// TIA Portal V19 export
FUNCTION_BLOCK "ALL_AI"   // FB3, FBD
{ S7_Optimized_Access := 'TRUE' }
// stored: MemoryReserve 100, SetENOAutomatically false
   VAR
      AI_TT01 { S7_SetPoint := 'True'} : "AI";
      AI_TT02 { S7_SetPoint := 'True'} : "AI";
      AI_TT03 { S7_SetPoint := 'True'} : "AI";
      AI_CHS_TT01 { S7_SetPoint := 'True'} : "AI";
      AI_CHS_TT02 { S7_SetPoint := 'True'} : "AI";
      AI_CHS_TT03 { S7_SetPoint := 'True'} : "AI";
      AI_CHS_TT04 { S7_SetPoint := 'True'} : "AI";
      AI_CHS_MGLT { S7_SetPoint := 'True'} : "AI";
      AI_R2_TT01 { S7_SetPoint := 'True'} : "AI";
      AI_R2_TT02 { S7_SetPoint := 'True'} : "AI";
      AI_R2_TT03 { S7_SetPoint := 'True'} : "AI";
      AI_R3_TT01 { S7_SetPoint := 'True'} : "AI";
      AI_R3_TT02 { S7_SetPoint := 'True'} : "AI";
      AI_R3_TT03 { S7_SetPoint := 'True'} : "AI";
      AI_R4_TT03 { S7_SetPoint := 'True'} : "AI";
      AI_R4_TT02 { S7_SetPoint := 'True'} : "AI";
      AI_R4_TT01 { S7_SetPoint := 'True'} : "AI";
      AI_R5_TT01 { S7_SetPoint := 'True'} : "AI";
      AI_R5_TT02 { S7_SetPoint := 'True'} : "AI";
      AI_R5_TT03 { S7_SetPoint := 'True'} : "AI";
      AI_R6_TT01 { S7_SetPoint := 'True'} : "AI";
      AI_R6_TT02 { S7_SetPoint := 'True'} : "AI";
      AI_R6_TT03 { S7_SetPoint := 'True'} : "AI";
      AI_R7_TT01 { S7_SetPoint := 'True'} : "AI";
      AI_R7_TT02 { S7_SetPoint := 'True'} : "AI";
      AI_R8_TT03 { S7_SetPoint := 'True'} : "AI";
      AI_R7_TT03 { S7_SetPoint := 'True'} : "AI";
      AI_R8_TT01 { S7_SetPoint := 'True'} : "AI";
      AI_R8_TT02 { S7_SetPoint := 'True'} : "AI";
      AI_R9_TT01 { S7_SetPoint := 'True'} : "AI";
      AI_R9_TT02 { S7_SetPoint := 'True'} : "AI";
      AI_R9_TT03 { S7_SetPoint := 'True'} : "AI";
      AI_R10_TT01 { S7_SetPoint := 'True'} : "AI";
      AI_R10_TT02 { S7_SetPoint := 'True'} : "AI";
      AI_R10_TT03 { S7_SetPoint := 'True'} : "AI";
      AI_R11_TT01 { S7_SetPoint := 'True'} : "AI";
      AI_R11_TT02 { S7_SetPoint := 'True'} : "AI";
      AI_R11_TT03 { S7_SetPoint := 'True'} : "AI";
      AI_R12_TT01 { S7_SetPoint := 'True'} : "AI";
      AI_R12_TT02 { S7_SetPoint := 'True'} : "AI";
      AI_R12_TT03 { S7_SetPoint := 'True'} : "AI";
      AI_R13_TT01 { S7_SetPoint := 'True'} : "AI";
      AI_R13_TT02 { S7_SetPoint := 'True'} : "AI";
      AI_R13_TT03 { S7_SetPoint := 'True'} : "AI";
      AI_R14_TT01 { S7_SetPoint := 'True'} : "AI";
      AI_R14_TT02 { S7_SetPoint := 'True'} : "AI";
      AI_R14_TT03 { S7_SetPoint := 'True'} : "AI";
      AI_R15_TT01 { S7_SetPoint := 'True'} : "AI";
      AI_R15_TT02 { S7_SetPoint := 'True'} : "AI";
      AI_R15_TT03 { S7_SetPoint := 'True'} : "AI";
      AI_R16_TT01 { S7_SetPoint := 'True'} : "AI";
      AI_R16_TT02 { S7_SetPoint := 'True'} : "AI";
      AI_R16_TT03 { S7_SetPoint := 'True'} : "AI";
      AI_R17_TT01 { S7_SetPoint := 'True'} : "AI";
      AI_R17_TT02 { S7_SetPoint := 'True'} : "AI";
      AI_R17_TT03 { S7_SetPoint := 'True'} : "AI";
      AI_R18_TT01 { S7_SetPoint := 'True'} : "AI";
      AI_R18_TT02 { S7_SetPoint := 'True'} : "AI";
      AI_R18_TT03 { S7_SetPoint := 'True'} : "AI";
      AI_CHS_PT { S7_SetPoint := 'True'} : "AI";
      AI_SMHS_TT01 { S7_SetPoint := 'True'} : "AI";
      AI_SMHS_TT02 { S7_SetPoint := 'True'} : "AI";
      AI_SMHS_TT03 { S7_SetPoint := 'True'} : "AI";
      AI_SMHS_TT04 { S7_SetPoint := 'True'} : "AI";
      AI_NMHS_TT01 { S7_SetPoint := 'True'} : "AI";
      AI_NMHS_TT02 { S7_SetPoint := 'True'} : "AI";
      AI_NMHS_TT03 { S7_SetPoint := 'True'} : "AI";
      AI_NMHS_TT04 { S7_SetPoint := 'True'} : "AI";
      AI_SMHS_PT01 { S7_SetPoint := 'True'} : "PT_AI";
      AI_SMHS_PT02 { S7_SetPoint := 'True'} : "PT_AI";
      AI_SMHS_PT03 { S7_SetPoint := 'True'} : "PT_AI";
      AI_SMHS_PT04 { S7_SetPoint := 'True'} : "PT_AI";
      AI_NMHS_PT04 { S7_SetPoint := 'True'} : "PT_AI";
      AI_NMHS_PT01 { S7_SetPoint := 'True'} : "PT_AI";
      AI_NMHS_PT02 { S7_SetPoint := 'True'} : "PT_AI";
      AI_NMHS_PT03 { S7_SetPoint := 'True'} : "PT_AI";
      AI_CS_TT01 { S7_SetPoint := 'True'} : "AI";
      AI_CS_TT02 { S7_SetPoint := 'True'} : "AI";
      AI_CS_TT03 { S7_SetPoint := 'True'} : "AI";
      AI_CS_TT04 { S7_SetPoint := 'True'} : "AI";
      AI_CS_MGLT { S7_SetPoint := 'True'} : "AI";
      AI_UCHS_TT01 { S7_SetPoint := 'True'} : "AI";
      AI_UCHS_TT02 { S7_SetPoint := 'True'} : "AI";
      AI_UCHS_TT03 { S7_SetPoint := 'True'} : "AI";
      AI_UCHS_TT04 { S7_SetPoint := 'True'} : "AI";
      AI_UCHS_MGLT { S7_SetPoint := 'True'} : "AI";
      AI_HS_TT01 { S7_SetPoint := 'True'} : "AI";
      AI_HS_TT02 { S7_SetPoint := 'True'} : "AI";
      AI_HS_TT03 { S7_SetPoint := 'True'} : "AI";
      AI_HS_MGLT { S7_SetPoint := 'True'} : "AI";
      "AI_A/SCRB_001_PH01" { S7_SetPoint := 'True'} : "AI";
      "AI_AI_A/SCRB_002_PH01" { S7_SetPoint := 'True'} : "AI";
      "AI_A/VP_01_APT01" { S7_SetPoint := 'True'} : "AI";
      "AI_A/VP_02_APT01" { S7_SetPoint := 'True'} : "AI";
      "AI_A/ANFD_001_APT01" { S7_SetPoint := 'True'} : "AI";
      "AI_A/ANFD_002_APT01" { S7_SetPoint := 'True'} : "AI";
      "AI_A/ANFD_003_APT01" { S7_SetPoint := 'True'} : "AI";
      AI_HS_TT9 { S7_SetPoint := 'True'} : "AI";
      "A/ANFD_001_TT01" { S7_SetPoint := 'True'} : "AI";
      "A/ANFD_002_TT01" { S7_SetPoint := 'True'} : "AI";
      "A/ANFD_003_TT01" { S7_SetPoint := 'True'} : "AI";
      "A/ANFD_004_TT01" { S7_SetPoint := 'True'} : "AI";
      AI_RCVD_001_APT01 { S7_SetPoint := 'True'} : "AI";
      AI_RCVD_002_APT01 { S7_SetPoint := 'True'} : "AI";
      AI_RCVD_001_TT01 { S7_SetPoint := 'True'} : "AI";
      AI_RCVD_002_TT01 { S7_SetPoint := 'True'} : "AI";
      "AI_A/VTD_001_APT01" { S7_SetPoint := 'True'} : "AI";
      "AI_A/VTD_002_APT01" { S7_SetPoint := 'True'} : "AI";
      "AI_A/VTD_001_TT01" { S7_SetPoint := 'True'} : "AI";
      "AI_A/VTD_002_TT01" { S7_SetPoint := 'True'} : "AI";
      "AI_A/TD_001_TT01" { S7_SetPoint := 'True'} : "AI";
      "AI_A/TD_002_TT01" { S7_SetPoint := 'True'} : "AI";
      DRIVE_RPM { S7_SetPoint := 'True'} : "DRIVE_RPM";
   END_VAR
BEGIN

REGION Network 1: ****REACTOR_1****
END_REGION

REGION Network 2: TT01
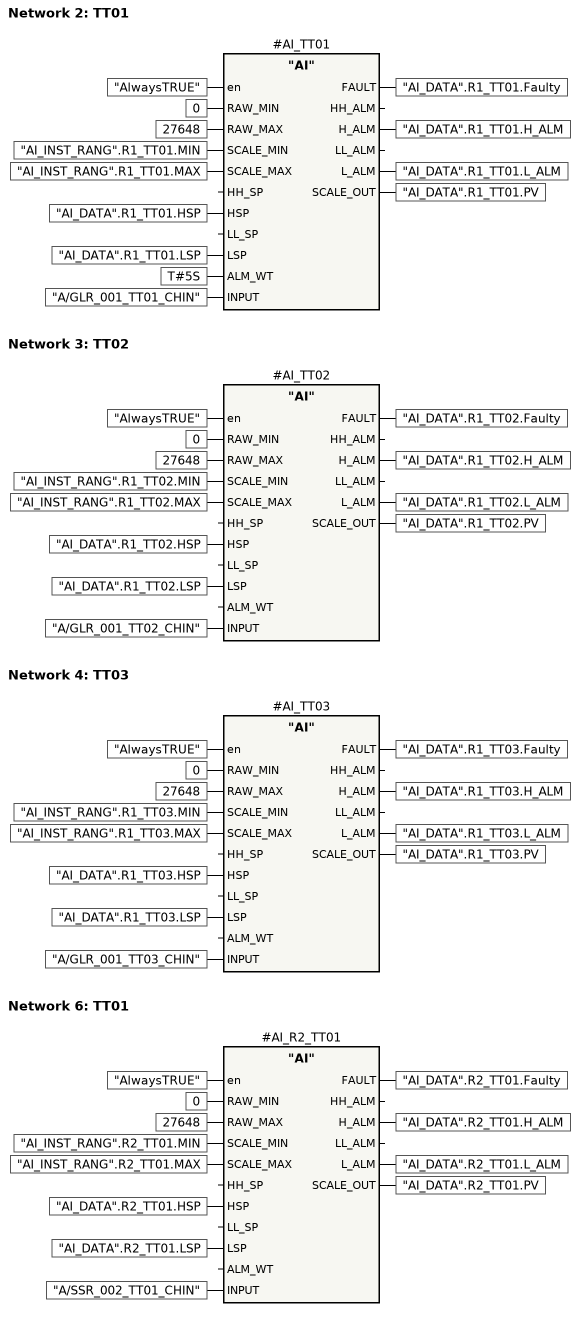
   IF "AlwaysTRUE" THEN
       #AI_TT01(RAW_MIN := 0,   // "AI"
                RAW_MAX := 27648,
                SCALE_MIN := "AI_INST_RANG".R1_TT01.MIN,
                SCALE_MAX := "AI_INST_RANG".R1_TT01.MAX,
                HSP := "AI_DATA".R1_TT01.HSP,
                LSP := "AI_DATA".R1_TT01.LSP,
                ALM_WT := T#5S,
                INPUT := "A/GLR_001_TT01_CHIN",
                FAULT => "AI_DATA".R1_TT01.Faulty,
                H_ALM => "AI_DATA".R1_TT01.H_ALM,
                L_ALM => "AI_DATA".R1_TT01.L_ALM,
                SCALE_OUT => "AI_DATA".R1_TT01.PV);
   END_IF;
END_REGION

REGION Network 3: TT02
   IF "AlwaysTRUE" THEN
       #AI_TT02(RAW_MIN := 0,   // "AI"
                RAW_MAX := 27648,
                SCALE_MIN := "AI_INST_RANG".R1_TT02.MIN,
                SCALE_MAX := "AI_INST_RANG".R1_TT02.MAX,
                HSP := "AI_DATA".R1_TT02.HSP,
                LSP := "AI_DATA".R1_TT02.LSP,
                INPUT := "A/GLR_001_TT02_CHIN",
                FAULT => "AI_DATA".R1_TT02.Faulty,
                H_ALM => "AI_DATA".R1_TT02.H_ALM,
                L_ALM => "AI_DATA".R1_TT02.L_ALM,
                SCALE_OUT => "AI_DATA".R1_TT02.PV);
   END_IF;
END_REGION

REGION Network 4: TT03
   IF "AlwaysTRUE" THEN
       #AI_TT03(RAW_MIN := 0,   // "AI"
                RAW_MAX := 27648,
                SCALE_MIN := "AI_INST_RANG".R1_TT03.MIN,
                SCALE_MAX := "AI_INST_RANG".R1_TT03.MAX,
                HSP := "AI_DATA".R1_TT03.HSP,
                LSP := "AI_DATA".R1_TT03.LSP,
                INPUT := "A/GLR_001_TT03_CHIN",
                FAULT => "AI_DATA".R1_TT03.Faulty,
                H_ALM => "AI_DATA".R1_TT03.H_ALM,
                L_ALM => "AI_DATA".R1_TT03.L_ALM,
                SCALE_OUT => "AI_DATA".R1_TT03.PV);
   END_IF;
END_REGION

REGION Network 5: ****REACTOR_2****
END_REGION

REGION Network 6: TT01
   IF "AlwaysTRUE" THEN
       #AI_R2_TT01(RAW_MIN := 0,   // "AI"
                   RAW_MAX := 27648,
                   SCALE_MIN := "AI_INST_RANG".R2_TT01.MIN,
                   SCALE_MAX := "AI_INST_RANG".R2_TT01.MAX,
                   HSP := "AI_DATA".R2_TT01.HSP,
                   LSP := "AI_DATA".R2_TT01.LSP,
                   INPUT := "A/SSR_002_TT01_CHIN",
                   FAULT => "AI_DATA".R2_TT01.Faulty,
                   H_ALM => "AI_DATA".R2_TT01.H_ALM,
                   L_ALM => "AI_DATA".R2_TT01.L_ALM,
                   SCALE_OUT => "AI_DATA".R2_TT01.PV);
   END_IF;
END_REGION

REGION Network 7: TT02
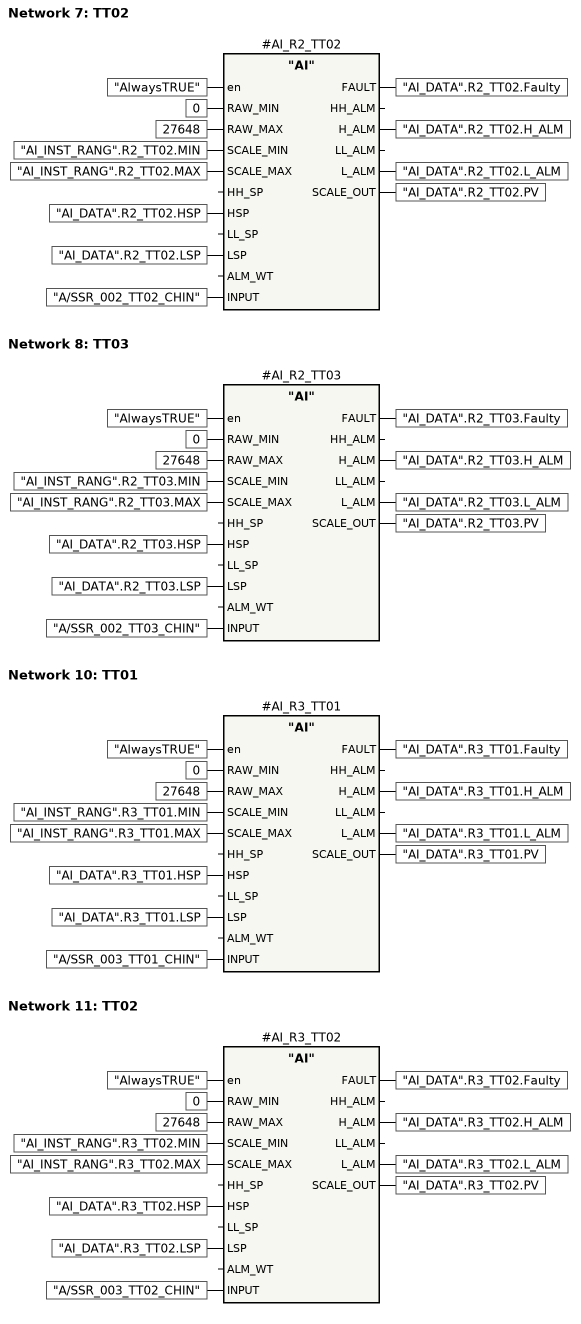
   IF "AlwaysTRUE" THEN
       #AI_R2_TT02(RAW_MIN := 0,   // "AI"
                   RAW_MAX := 27648,
                   SCALE_MIN := "AI_INST_RANG".R2_TT02.MIN,
                   SCALE_MAX := "AI_INST_RANG".R2_TT02.MAX,
                   HSP := "AI_DATA".R2_TT02.HSP,
                   LSP := "AI_DATA".R2_TT02.LSP,
                   INPUT := "A/SSR_002_TT02_CHIN",
                   FAULT => "AI_DATA".R2_TT02.Faulty,
                   H_ALM => "AI_DATA".R2_TT02.H_ALM,
                   L_ALM => "AI_DATA".R2_TT02.L_ALM,
                   SCALE_OUT => "AI_DATA".R2_TT02.PV);
   END_IF;
END_REGION

REGION Network 8: TT03
   IF "AlwaysTRUE" THEN
       #AI_R2_TT03(RAW_MIN := 0,   // "AI"
                   RAW_MAX := 27648,
                   SCALE_MIN := "AI_INST_RANG".R2_TT03.MIN,
                   SCALE_MAX := "AI_INST_RANG".R2_TT03.MAX,
                   HSP := "AI_DATA".R2_TT03.HSP,
                   LSP := "AI_DATA".R2_TT03.LSP,
                   INPUT := "A/SSR_002_TT03_CHIN",
                   FAULT => "AI_DATA".R2_TT03.Faulty,
                   H_ALM => "AI_DATA".R2_TT03.H_ALM,
                   L_ALM => "AI_DATA".R2_TT03.L_ALM,
                   SCALE_OUT => "AI_DATA".R2_TT03.PV);
   END_IF;
END_REGION

REGION Network 9: ****REACTOR_3****
END_REGION

REGION Network 10: TT01
   IF "AlwaysTRUE" THEN
       #AI_R3_TT01(RAW_MIN := 0,   // "AI"
                   RAW_MAX := 27648,
                   SCALE_MIN := "AI_INST_RANG".R3_TT01.MIN,
                   SCALE_MAX := "AI_INST_RANG".R3_TT01.MAX,
                   HSP := "AI_DATA".R3_TT01.HSP,
                   LSP := "AI_DATA".R3_TT01.LSP,
                   INPUT := "A/SSR_003_TT01_CHIN",
                   FAULT => "AI_DATA".R3_TT01.Faulty,
                   H_ALM => "AI_DATA".R3_TT01.H_ALM,
                   L_ALM => "AI_DATA".R3_TT01.L_ALM,
                   SCALE_OUT => "AI_DATA".R3_TT01.PV);
   END_IF;
END_REGION

REGION Network 11: TT02
   IF "AlwaysTRUE" THEN
       #AI_R3_TT02(RAW_MIN := 0,   // "AI"
                   RAW_MAX := 27648,
                   SCALE_MIN := "AI_INST_RANG".R3_TT02.MIN,
                   SCALE_MAX := "AI_INST_RANG".R3_TT02.MAX,
                   HSP := "AI_DATA".R3_TT02.HSP,
                   LSP := "AI_DATA".R3_TT02.LSP,
                   INPUT := "A/SSR_003_TT02_CHIN",
                   FAULT => "AI_DATA".R3_TT02.Faulty,
                   H_ALM => "AI_DATA".R3_TT02.H_ALM,
                   L_ALM => "AI_DATA".R3_TT02.L_ALM,
                   SCALE_OUT => "AI_DATA".R3_TT02.PV);
   END_IF;
END_REGION

REGION Network 12: TT03
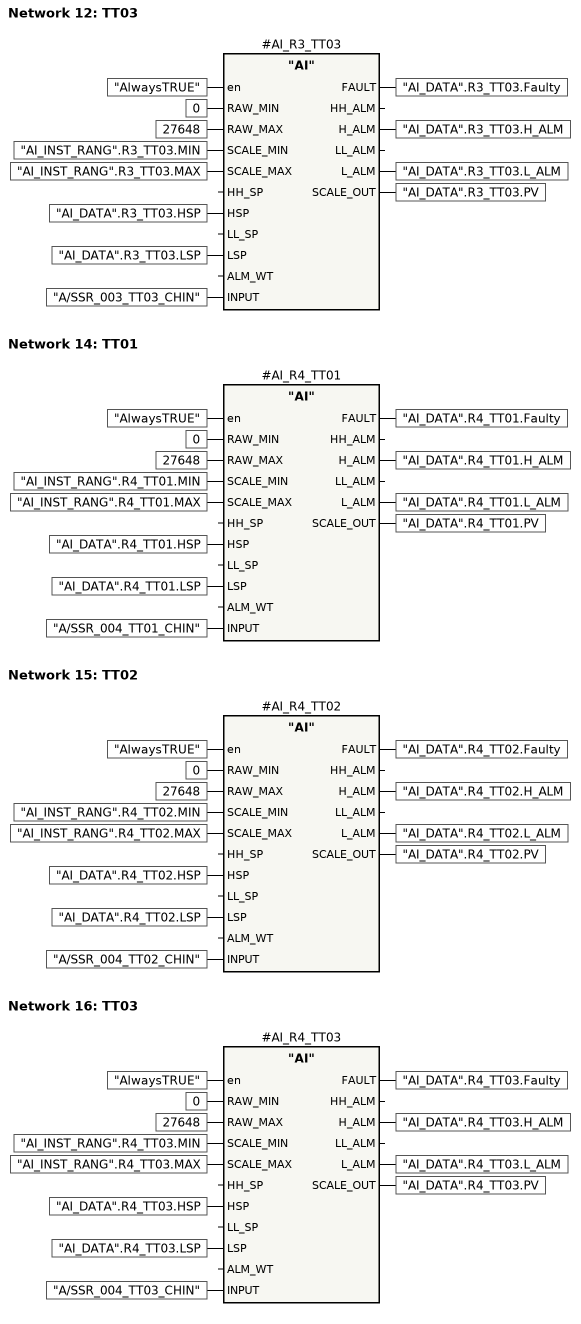
   IF "AlwaysTRUE" THEN
       #AI_R3_TT03(RAW_MIN := 0,   // "AI"
                   RAW_MAX := 27648,
                   SCALE_MIN := "AI_INST_RANG".R3_TT03.MIN,
                   SCALE_MAX := "AI_INST_RANG".R3_TT03.MAX,
                   HSP := "AI_DATA".R3_TT03.HSP,
                   LSP := "AI_DATA".R3_TT03.LSP,
                   INPUT := "A/SSR_003_TT03_CHIN",
                   FAULT => "AI_DATA".R3_TT03.Faulty,
                   H_ALM => "AI_DATA".R3_TT03.H_ALM,
                   L_ALM => "AI_DATA".R3_TT03.L_ALM,
                   SCALE_OUT => "AI_DATA".R3_TT03.PV);
   END_IF;
END_REGION

REGION Network 13: ****REACTOR_4****
END_REGION

REGION Network 14: TT01
   IF "AlwaysTRUE" THEN
       #AI_R4_TT01(RAW_MIN := 0,   // "AI"
                   RAW_MAX := 27648,
                   SCALE_MIN := "AI_INST_RANG".R4_TT01.MIN,
                   SCALE_MAX := "AI_INST_RANG".R4_TT01.MAX,
                   HSP := "AI_DATA".R4_TT01.HSP,
                   LSP := "AI_DATA".R4_TT01.LSP,
                   INPUT := "A/SSR_004_TT01_CHIN",
                   FAULT => "AI_DATA".R4_TT01.Faulty,
                   H_ALM => "AI_DATA".R4_TT01.H_ALM,
                   L_ALM => "AI_DATA".R4_TT01.L_ALM,
                   SCALE_OUT => "AI_DATA".R4_TT01.PV);
   END_IF;
END_REGION

REGION Network 15: TT02
   IF "AlwaysTRUE" THEN
       #AI_R4_TT02(RAW_MIN := 0,   // "AI"
                   RAW_MAX := 27648,
                   SCALE_MIN := "AI_INST_RANG".R4_TT02.MIN,
                   SCALE_MAX := "AI_INST_RANG".R4_TT02.MAX,
                   HSP := "AI_DATA".R4_TT02.HSP,
                   LSP := "AI_DATA".R4_TT02.LSP,
                   INPUT := "A/SSR_004_TT02_CHIN",
                   FAULT => "AI_DATA".R4_TT02.Faulty,
                   H_ALM => "AI_DATA".R4_TT02.H_ALM,
                   L_ALM => "AI_DATA".R4_TT02.L_ALM,
                   SCALE_OUT => "AI_DATA".R4_TT02.PV);
   END_IF;
END_REGION

REGION Network 16: TT03
   IF "AlwaysTRUE" THEN
       #AI_R4_TT03(RAW_MIN := 0,   // "AI"
                   RAW_MAX := 27648,
                   SCALE_MIN := "AI_INST_RANG".R4_TT03.MIN,
                   SCALE_MAX := "AI_INST_RANG".R4_TT03.MAX,
                   HSP := "AI_DATA".R4_TT03.HSP,
                   LSP := "AI_DATA".R4_TT03.LSP,
                   INPUT := "A/SSR_004_TT03_CHIN",
                   FAULT => "AI_DATA".R4_TT03.Faulty,
                   H_ALM => "AI_DATA".R4_TT03.H_ALM,
                   L_ALM => "AI_DATA".R4_TT03.L_ALM,
                   SCALE_OUT => "AI_DATA".R4_TT03.PV);
   END_IF;
END_REGION

REGION Network 17: ****REACTOR_5****
END_REGION

REGION Network 18: TT01
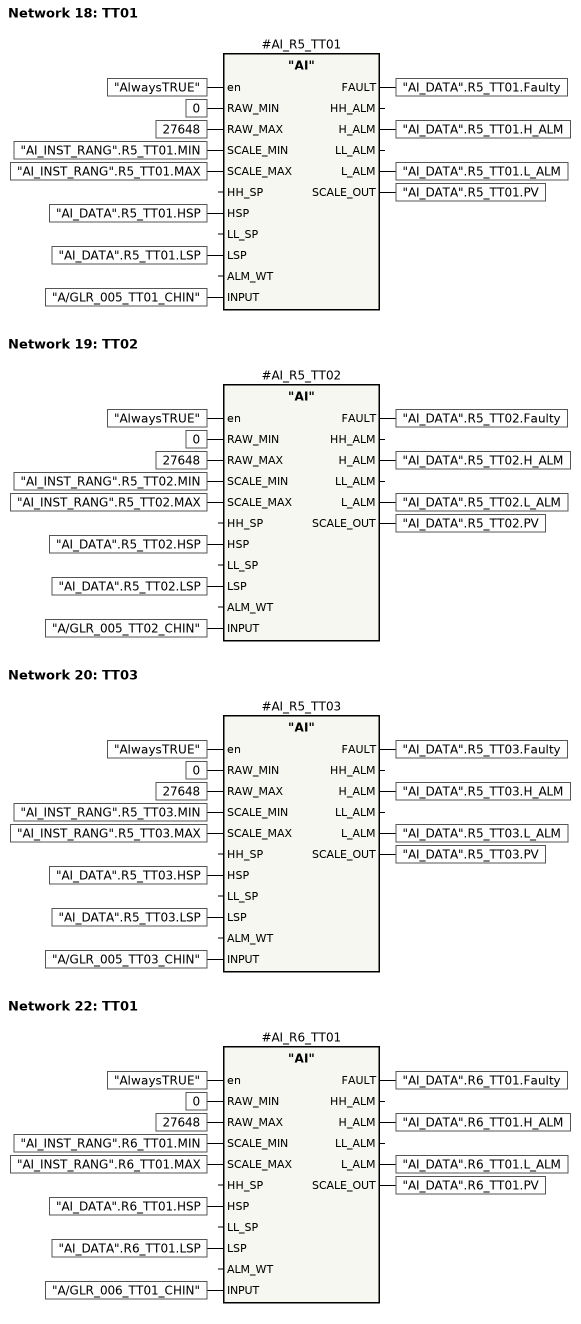
   IF "AlwaysTRUE" THEN
       #AI_R5_TT01(RAW_MIN := 0,   // "AI"
                   RAW_MAX := 27648,
                   SCALE_MIN := "AI_INST_RANG".R5_TT01.MIN,
                   SCALE_MAX := "AI_INST_RANG".R5_TT01.MAX,
                   HSP := "AI_DATA".R5_TT01.HSP,
                   LSP := "AI_DATA".R5_TT01.LSP,
                   INPUT := "A/GLR_005_TT01_CHIN",
                   FAULT => "AI_DATA".R5_TT01.Faulty,
                   H_ALM => "AI_DATA".R5_TT01.H_ALM,
                   L_ALM => "AI_DATA".R5_TT01.L_ALM,
                   SCALE_OUT => "AI_DATA".R5_TT01.PV);
   END_IF;
END_REGION

REGION Network 19: TT02
   IF "AlwaysTRUE" THEN
       #AI_R5_TT02(RAW_MIN := 0,   // "AI"
                   RAW_MAX := 27648,
                   SCALE_MIN := "AI_INST_RANG".R5_TT02.MIN,
                   SCALE_MAX := "AI_INST_RANG".R5_TT02.MAX,
                   HSP := "AI_DATA".R5_TT02.HSP,
                   LSP := "AI_DATA".R5_TT02.LSP,
                   INPUT := "A/GLR_005_TT02_CHIN",
                   FAULT => "AI_DATA".R5_TT02.Faulty,
                   H_ALM => "AI_DATA".R5_TT02.H_ALM,
                   L_ALM => "AI_DATA".R5_TT02.L_ALM,
                   SCALE_OUT => "AI_DATA".R5_TT02.PV);
   END_IF;
END_REGION

REGION Network 20: TT03
   IF "AlwaysTRUE" THEN
       #AI_R5_TT03(RAW_MIN := 0,   // "AI"
                   RAW_MAX := 27648,
                   SCALE_MIN := "AI_INST_RANG".R5_TT03.MIN,
                   SCALE_MAX := "AI_INST_RANG".R5_TT03.MAX,
                   HSP := "AI_DATA".R5_TT03.HSP,
                   LSP := "AI_DATA".R5_TT03.LSP,
                   INPUT := "A/GLR_005_TT03_CHIN",
                   FAULT => "AI_DATA".R5_TT03.Faulty,
                   H_ALM => "AI_DATA".R5_TT03.H_ALM,
                   L_ALM => "AI_DATA".R5_TT03.L_ALM,
                   SCALE_OUT => "AI_DATA".R5_TT03.PV);
   END_IF;
END_REGION

REGION Network 21: ****REACTOR_6****
END_REGION

REGION Network 22: TT01
   IF "AlwaysTRUE" THEN
       #AI_R6_TT01(RAW_MIN := 0,   // "AI"
                   RAW_MAX := 27648,
                   SCALE_MIN := "AI_INST_RANG".R6_TT01.MIN,
                   SCALE_MAX := "AI_INST_RANG".R6_TT01.MAX,
                   HSP := "AI_DATA".R6_TT01.HSP,
                   LSP := "AI_DATA".R6_TT01.LSP,
                   INPUT := "A/GLR_006_TT01_CHIN",
                   FAULT => "AI_DATA".R6_TT01.Faulty,
                   H_ALM => "AI_DATA".R6_TT01.H_ALM,
                   L_ALM => "AI_DATA".R6_TT01.L_ALM,
                   SCALE_OUT => "AI_DATA".R6_TT01.PV);
   END_IF;
END_REGION

REGION Network 23: TT02
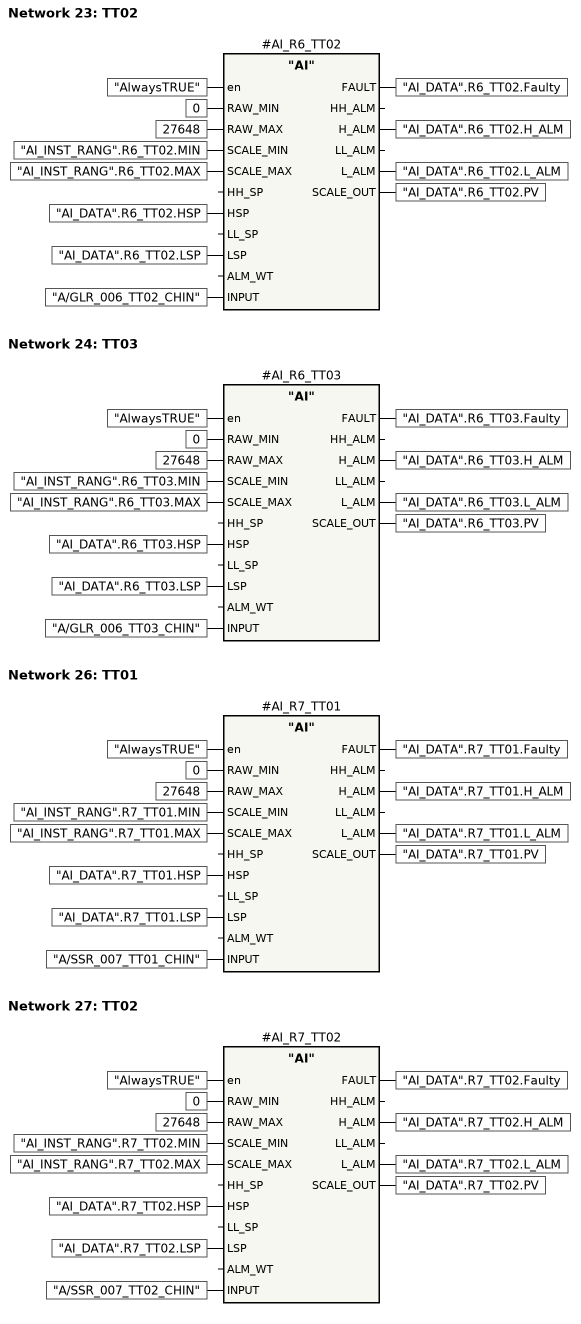
   IF "AlwaysTRUE" THEN
       #AI_R6_TT02(RAW_MIN := 0,   // "AI"
                   RAW_MAX := 27648,
                   SCALE_MIN := "AI_INST_RANG".R6_TT02.MIN,
                   SCALE_MAX := "AI_INST_RANG".R6_TT02.MAX,
                   HSP := "AI_DATA".R6_TT02.HSP,
                   LSP := "AI_DATA".R6_TT02.LSP,
                   INPUT := "A/GLR_006_TT02_CHIN",
                   FAULT => "AI_DATA".R6_TT02.Faulty,
                   H_ALM => "AI_DATA".R6_TT02.H_ALM,
                   L_ALM => "AI_DATA".R6_TT02.L_ALM,
                   SCALE_OUT => "AI_DATA".R6_TT02.PV);
   END_IF;
END_REGION

REGION Network 24: TT03
   IF "AlwaysTRUE" THEN
       #AI_R6_TT03(RAW_MIN := 0,   // "AI"
                   RAW_MAX := 27648,
                   SCALE_MIN := "AI_INST_RANG".R6_TT03.MIN,
                   SCALE_MAX := "AI_INST_RANG".R6_TT03.MAX,
                   HSP := "AI_DATA".R6_TT03.HSP,
                   LSP := "AI_DATA".R6_TT03.LSP,
                   INPUT := "A/GLR_006_TT03_CHIN",
                   FAULT => "AI_DATA".R6_TT03.Faulty,
                   H_ALM => "AI_DATA".R6_TT03.H_ALM,
                   L_ALM => "AI_DATA".R6_TT03.L_ALM,
                   SCALE_OUT => "AI_DATA".R6_TT03.PV);
   END_IF;
END_REGION

REGION Network 25: ****REACTOR_7****
END_REGION

REGION Network 26: TT01
   IF "AlwaysTRUE" THEN
       #AI_R7_TT01(RAW_MIN := 0,   // "AI"
                   RAW_MAX := 27648,
                   SCALE_MIN := "AI_INST_RANG".R7_TT01.MIN,
                   SCALE_MAX := "AI_INST_RANG".R7_TT01.MAX,
                   HSP := "AI_DATA".R7_TT01.HSP,
                   LSP := "AI_DATA".R7_TT01.LSP,
                   INPUT := "A/SSR_007_TT01_CHIN",
                   FAULT => "AI_DATA".R7_TT01.Faulty,
                   H_ALM => "AI_DATA".R7_TT01.H_ALM,
                   L_ALM => "AI_DATA".R7_TT01.L_ALM,
                   SCALE_OUT => "AI_DATA".R7_TT01.PV);
   END_IF;
END_REGION

REGION Network 27: TT02
   IF "AlwaysTRUE" THEN
       #AI_R7_TT02(RAW_MIN := 0,   // "AI"
                   RAW_MAX := 27648,
                   SCALE_MIN := "AI_INST_RANG".R7_TT02.MIN,
                   SCALE_MAX := "AI_INST_RANG".R7_TT02.MAX,
                   HSP := "AI_DATA".R7_TT02.HSP,
                   LSP := "AI_DATA".R7_TT02.LSP,
                   INPUT := "A/SSR_007_TT02_CHIN",
                   FAULT => "AI_DATA".R7_TT02.Faulty,
                   H_ALM => "AI_DATA".R7_TT02.H_ALM,
                   L_ALM => "AI_DATA".R7_TT02.L_ALM,
                   SCALE_OUT => "AI_DATA".R7_TT02.PV);
   END_IF;
END_REGION

REGION Network 28: TT03
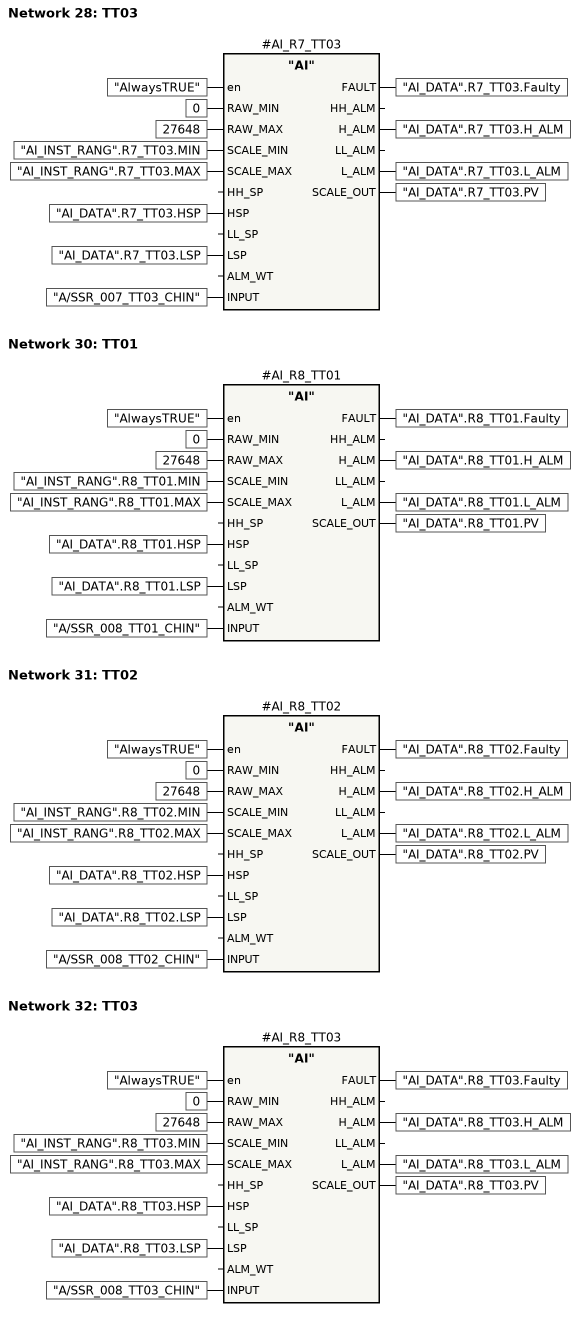
   IF "AlwaysTRUE" THEN
       #AI_R7_TT03(RAW_MIN := 0,   // "AI"
                   RAW_MAX := 27648,
                   SCALE_MIN := "AI_INST_RANG".R7_TT03.MIN,
                   SCALE_MAX := "AI_INST_RANG".R7_TT03.MAX,
                   HSP := "AI_DATA".R7_TT03.HSP,
                   LSP := "AI_DATA".R7_TT03.LSP,
                   INPUT := "A/SSR_007_TT03_CHIN",
                   FAULT => "AI_DATA".R7_TT03.Faulty,
                   H_ALM => "AI_DATA".R7_TT03.H_ALM,
                   L_ALM => "AI_DATA".R7_TT03.L_ALM,
                   SCALE_OUT => "AI_DATA".R7_TT03.PV);
   END_IF;
END_REGION

REGION Network 29: ****REACTOR_8****
END_REGION

REGION Network 30: TT01
   IF "AlwaysTRUE" THEN
       #AI_R8_TT01(RAW_MIN := 0,   // "AI"
                   RAW_MAX := 27648,
                   SCALE_MIN := "AI_INST_RANG".R8_TT01.MIN,
                   SCALE_MAX := "AI_INST_RANG".R8_TT01.MAX,
                   HSP := "AI_DATA".R8_TT01.HSP,
                   LSP := "AI_DATA".R8_TT01.LSP,
                   INPUT := "A/SSR_008_TT01_CHIN",
                   FAULT => "AI_DATA".R8_TT01.Faulty,
                   H_ALM => "AI_DATA".R8_TT01.H_ALM,
                   L_ALM => "AI_DATA".R8_TT01.L_ALM,
                   SCALE_OUT => "AI_DATA".R8_TT01.PV);
   END_IF;
END_REGION

REGION Network 31: TT02
   IF "AlwaysTRUE" THEN
       #AI_R8_TT02(RAW_MIN := 0,   // "AI"
                   RAW_MAX := 27648,
                   SCALE_MIN := "AI_INST_RANG".R8_TT02.MIN,
                   SCALE_MAX := "AI_INST_RANG".R8_TT02.MAX,
                   HSP := "AI_DATA".R8_TT02.HSP,
                   LSP := "AI_DATA".R8_TT02.LSP,
                   INPUT := "A/SSR_008_TT02_CHIN",
                   FAULT => "AI_DATA".R8_TT02.Faulty,
                   H_ALM => "AI_DATA".R8_TT02.H_ALM,
                   L_ALM => "AI_DATA".R8_TT02.L_ALM,
                   SCALE_OUT => "AI_DATA".R8_TT02.PV);
   END_IF;
END_REGION

REGION Network 32: TT03
   IF "AlwaysTRUE" THEN
       #AI_R8_TT03(RAW_MIN := 0,   // "AI"
                   RAW_MAX := 27648,
                   SCALE_MIN := "AI_INST_RANG".R8_TT03.MIN,
                   SCALE_MAX := "AI_INST_RANG".R8_TT03.MAX,
                   HSP := "AI_DATA".R8_TT03.HSP,
                   LSP := "AI_DATA".R8_TT03.LSP,
                   INPUT := "A/SSR_008_TT03_CHIN",
                   FAULT => "AI_DATA".R8_TT03.Faulty,
                   H_ALM => "AI_DATA".R8_TT03.H_ALM,
                   L_ALM => "AI_DATA".R8_TT03.L_ALM,
                   SCALE_OUT => "AI_DATA".R8_TT03.PV);
   END_IF;
END_REGION

REGION Network 33: ****REACTOR_9****
END_REGION

REGION Network 34: TT01
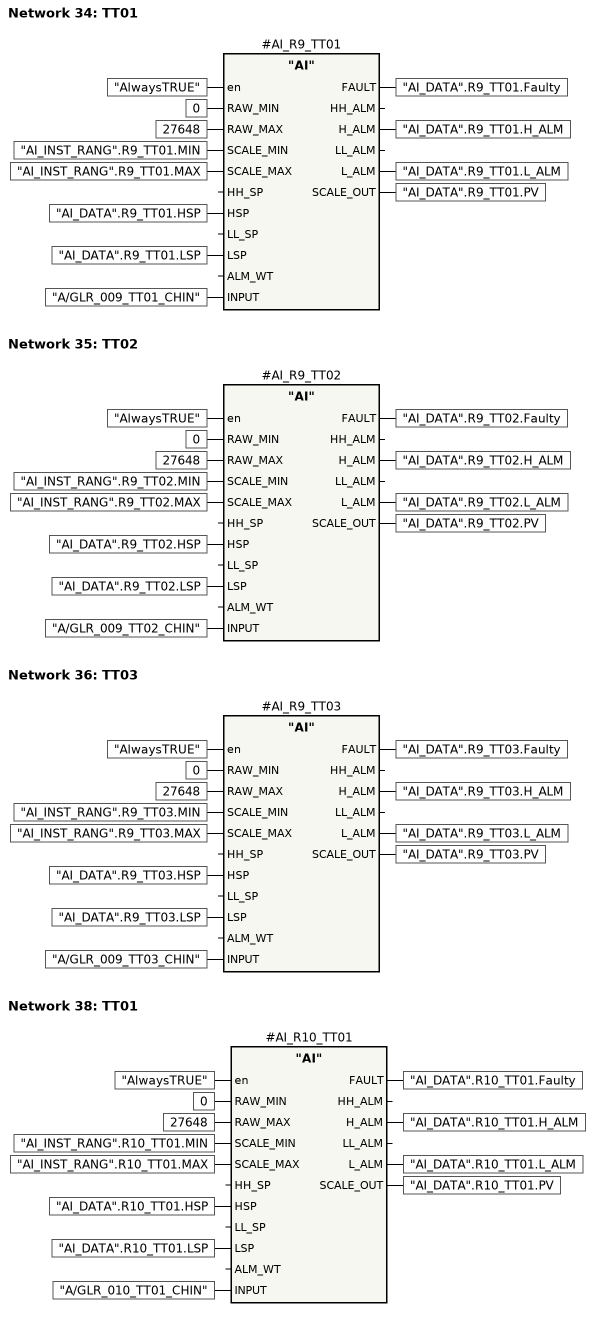
   IF "AlwaysTRUE" THEN
       #AI_R9_TT01(RAW_MIN := 0,   // "AI"
                   RAW_MAX := 27648,
                   SCALE_MIN := "AI_INST_RANG".R9_TT01.MIN,
                   SCALE_MAX := "AI_INST_RANG".R9_TT01.MAX,
                   HSP := "AI_DATA".R9_TT01.HSP,
                   LSP := "AI_DATA".R9_TT01.LSP,
                   INPUT := "A/GLR_009_TT01_CHIN",
                   FAULT => "AI_DATA".R9_TT01.Faulty,
                   H_ALM => "AI_DATA".R9_TT01.H_ALM,
                   L_ALM => "AI_DATA".R9_TT01.L_ALM,
                   SCALE_OUT => "AI_DATA".R9_TT01.PV);
   END_IF;
END_REGION

REGION Network 35: TT02
   IF "AlwaysTRUE" THEN
       #AI_R9_TT02(RAW_MIN := 0,   // "AI"
                   RAW_MAX := 27648,
                   SCALE_MIN := "AI_INST_RANG".R9_TT02.MIN,
                   SCALE_MAX := "AI_INST_RANG".R9_TT02.MAX,
                   HSP := "AI_DATA".R9_TT02.HSP,
                   LSP := "AI_DATA".R9_TT02.LSP,
                   INPUT := "A/GLR_009_TT02_CHIN",
                   FAULT => "AI_DATA".R9_TT02.Faulty,
                   H_ALM => "AI_DATA".R9_TT02.H_ALM,
                   L_ALM => "AI_DATA".R9_TT02.L_ALM,
                   SCALE_OUT => "AI_DATA".R9_TT02.PV);
   END_IF;
END_REGION

REGION Network 36: TT03
   IF "AlwaysTRUE" THEN
       #AI_R9_TT03(RAW_MIN := 0,   // "AI"
                   RAW_MAX := 27648,
                   SCALE_MIN := "AI_INST_RANG".R9_TT03.MIN,
                   SCALE_MAX := "AI_INST_RANG".R9_TT03.MAX,
                   HSP := "AI_DATA".R9_TT03.HSP,
                   LSP := "AI_DATA".R9_TT03.LSP,
                   INPUT := "A/GLR_009_TT03_CHIN",
                   FAULT => "AI_DATA".R9_TT03.Faulty,
                   H_ALM => "AI_DATA".R9_TT03.H_ALM,
                   L_ALM => "AI_DATA".R9_TT03.L_ALM,
                   SCALE_OUT => "AI_DATA".R9_TT03.PV);
   END_IF;
END_REGION

REGION Network 37: ****REACTOR_10****
END_REGION

REGION Network 38: TT01
   IF "AlwaysTRUE" THEN
       #AI_R10_TT01(RAW_MIN := 0,   // "AI"
                    RAW_MAX := 27648,
                    SCALE_MIN := "AI_INST_RANG".R10_TT01.MIN,
                    SCALE_MAX := "AI_INST_RANG".R10_TT01.MAX,
                    HSP := "AI_DATA".R10_TT01.HSP,
                    LSP := "AI_DATA".R10_TT01.LSP,
                    INPUT := "A/GLR_010_TT01_CHIN",
                    FAULT => "AI_DATA".R10_TT01.Faulty,
                    H_ALM => "AI_DATA".R10_TT01.H_ALM,
                    L_ALM => "AI_DATA".R10_TT01.L_ALM,
                    SCALE_OUT => "AI_DATA".R10_TT01.PV);
   END_IF;
END_REGION

REGION Network 39: TT02
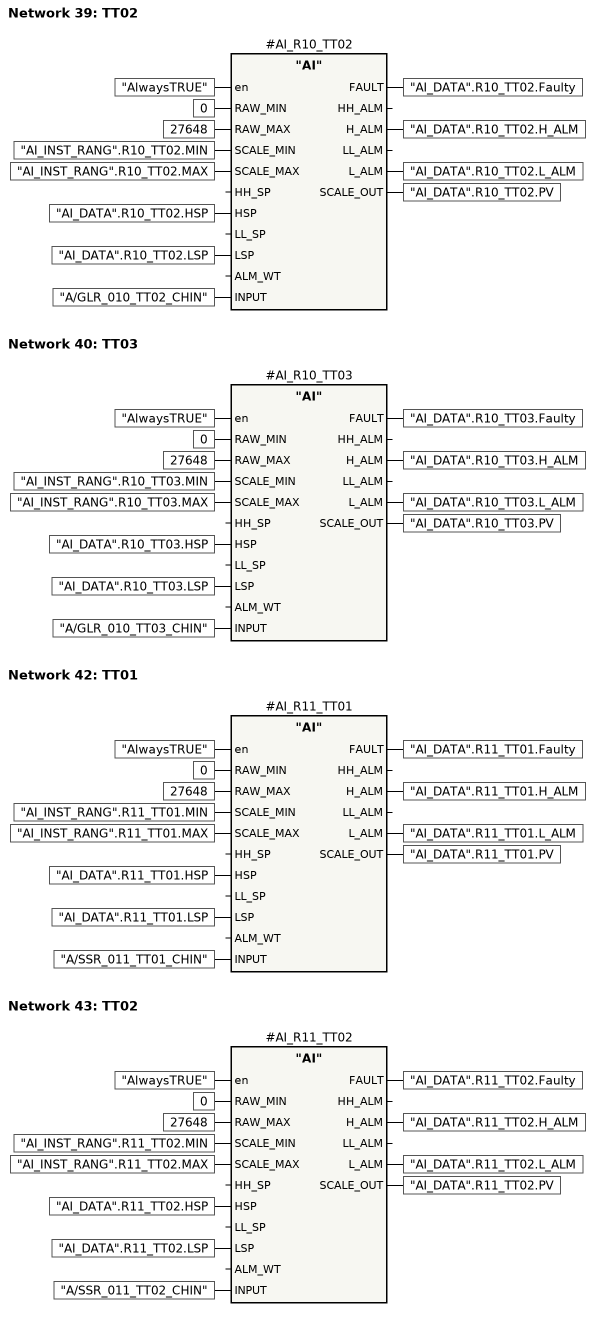
   IF "AlwaysTRUE" THEN
       #AI_R10_TT02(RAW_MIN := 0,   // "AI"
                    RAW_MAX := 27648,
                    SCALE_MIN := "AI_INST_RANG".R10_TT02.MIN,
                    SCALE_MAX := "AI_INST_RANG".R10_TT02.MAX,
                    HSP := "AI_DATA".R10_TT02.HSP,
                    LSP := "AI_DATA".R10_TT02.LSP,
                    INPUT := "A/GLR_010_TT02_CHIN",
                    FAULT => "AI_DATA".R10_TT02.Faulty,
                    H_ALM => "AI_DATA".R10_TT02.H_ALM,
                    L_ALM => "AI_DATA".R10_TT02.L_ALM,
                    SCALE_OUT => "AI_DATA".R10_TT02.PV);
   END_IF;
END_REGION

REGION Network 40: TT03
   IF "AlwaysTRUE" THEN
       #AI_R10_TT03(RAW_MIN := 0,   // "AI"
                    RAW_MAX := 27648,
                    SCALE_MIN := "AI_INST_RANG".R10_TT03.MIN,
                    SCALE_MAX := "AI_INST_RANG".R10_TT03.MAX,
                    HSP := "AI_DATA".R10_TT03.HSP,
                    LSP := "AI_DATA".R10_TT03.LSP,
                    INPUT := "A/GLR_010_TT03_CHIN",
                    FAULT => "AI_DATA".R10_TT03.Faulty,
                    H_ALM => "AI_DATA".R10_TT03.H_ALM,
                    L_ALM => "AI_DATA".R10_TT03.L_ALM,
                    SCALE_OUT => "AI_DATA".R10_TT03.PV);
   END_IF;
END_REGION

REGION Network 41: ****REACTOR_11****
END_REGION

REGION Network 42: TT01
   IF "AlwaysTRUE" THEN
       #AI_R11_TT01(RAW_MIN := 0,   // "AI"
                    RAW_MAX := 27648,
                    SCALE_MIN := "AI_INST_RANG".R11_TT01.MIN,
                    SCALE_MAX := "AI_INST_RANG".R11_TT01.MAX,
                    HSP := "AI_DATA".R11_TT01.HSP,
                    LSP := "AI_DATA".R11_TT01.LSP,
                    INPUT := "A/SSR_011_TT01_CHIN",
                    FAULT => "AI_DATA".R11_TT01.Faulty,
                    H_ALM => "AI_DATA".R11_TT01.H_ALM,
                    L_ALM => "AI_DATA".R11_TT01.L_ALM,
                    SCALE_OUT => "AI_DATA".R11_TT01.PV);
   END_IF;
END_REGION

REGION Network 43: TT02
   IF "AlwaysTRUE" THEN
       #AI_R11_TT02(RAW_MIN := 0,   // "AI"
                    RAW_MAX := 27648,
                    SCALE_MIN := "AI_INST_RANG".R11_TT02.MIN,
                    SCALE_MAX := "AI_INST_RANG".R11_TT02.MAX,
                    HSP := "AI_DATA".R11_TT02.HSP,
                    LSP := "AI_DATA".R11_TT02.LSP,
                    INPUT := "A/SSR_011_TT02_CHIN",
                    FAULT => "AI_DATA".R11_TT02.Faulty,
                    H_ALM => "AI_DATA".R11_TT02.H_ALM,
                    L_ALM => "AI_DATA".R11_TT02.L_ALM,
                    SCALE_OUT => "AI_DATA".R11_TT02.PV);
   END_IF;
END_REGION

REGION Network 44: TT03
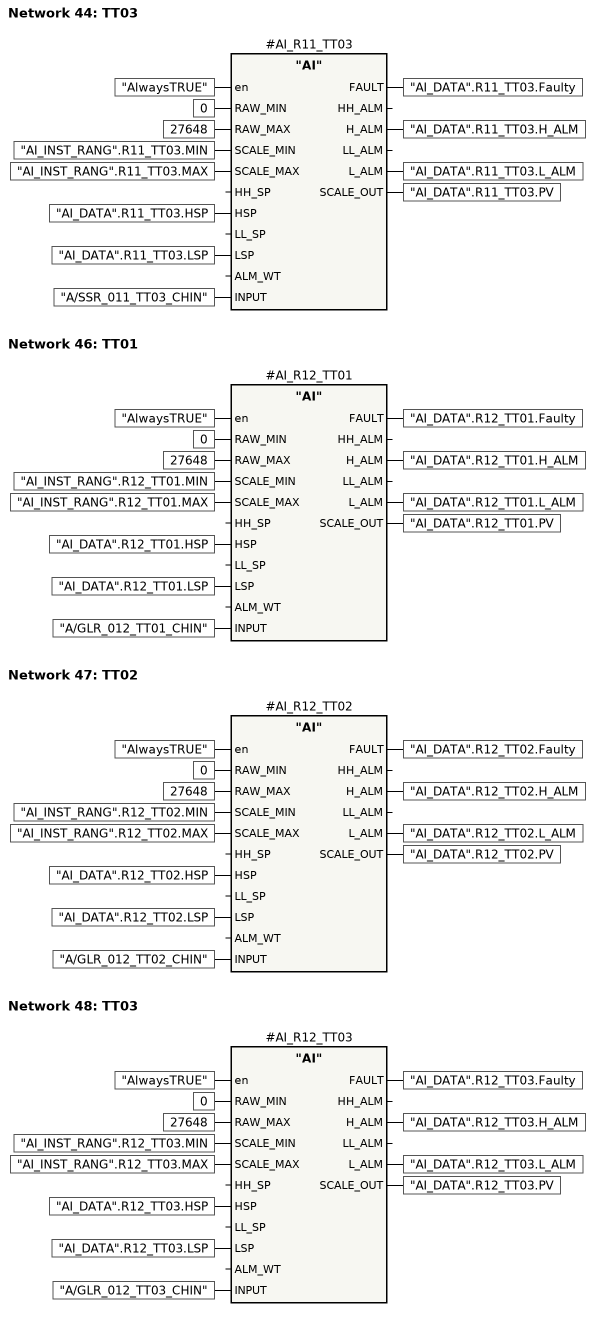
   IF "AlwaysTRUE" THEN
       #AI_R11_TT03(RAW_MIN := 0,   // "AI"
                    RAW_MAX := 27648,
                    SCALE_MIN := "AI_INST_RANG".R11_TT03.MIN,
                    SCALE_MAX := "AI_INST_RANG".R11_TT03.MAX,
                    HSP := "AI_DATA".R11_TT03.HSP,
                    LSP := "AI_DATA".R11_TT03.LSP,
                    INPUT := "A/SSR_011_TT03_CHIN",
                    FAULT => "AI_DATA".R11_TT03.Faulty,
                    H_ALM => "AI_DATA".R11_TT03.H_ALM,
                    L_ALM => "AI_DATA".R11_TT03.L_ALM,
                    SCALE_OUT => "AI_DATA".R11_TT03.PV);
   END_IF;
END_REGION

REGION Network 45: ****REACTOR_12****
END_REGION

REGION Network 46: TT01
   IF "AlwaysTRUE" THEN
       #AI_R12_TT01(RAW_MIN := 0,   // "AI"
                    RAW_MAX := 27648,
                    SCALE_MIN := "AI_INST_RANG".R12_TT01.MIN,
                    SCALE_MAX := "AI_INST_RANG".R12_TT01.MAX,
                    HSP := "AI_DATA".R12_TT01.HSP,
                    LSP := "AI_DATA".R12_TT01.LSP,
                    INPUT := "A/GLR_012_TT01_CHIN",
                    FAULT => "AI_DATA".R12_TT01.Faulty,
                    H_ALM => "AI_DATA".R12_TT01.H_ALM,
                    L_ALM => "AI_DATA".R12_TT01.L_ALM,
                    SCALE_OUT => "AI_DATA".R12_TT01.PV);
   END_IF;
END_REGION

REGION Network 47: TT02
   IF "AlwaysTRUE" THEN
       #AI_R12_TT02(RAW_MIN := 0,   // "AI"
                    RAW_MAX := 27648,
                    SCALE_MIN := "AI_INST_RANG".R12_TT02.MIN,
                    SCALE_MAX := "AI_INST_RANG".R12_TT02.MAX,
                    HSP := "AI_DATA".R12_TT02.HSP,
                    LSP := "AI_DATA".R12_TT02.LSP,
                    INPUT := "A/GLR_012_TT02_CHIN",
                    FAULT => "AI_DATA".R12_TT02.Faulty,
                    H_ALM => "AI_DATA".R12_TT02.H_ALM,
                    L_ALM => "AI_DATA".R12_TT02.L_ALM,
                    SCALE_OUT => "AI_DATA".R12_TT02.PV);
   END_IF;
END_REGION

REGION Network 48: TT03
   IF "AlwaysTRUE" THEN
       #AI_R12_TT03(RAW_MIN := 0,   // "AI"
                    RAW_MAX := 27648,
                    SCALE_MIN := "AI_INST_RANG".R12_TT03.MIN,
                    SCALE_MAX := "AI_INST_RANG".R12_TT03.MAX,
                    HSP := "AI_DATA".R12_TT03.HSP,
                    LSP := "AI_DATA".R12_TT03.LSP,
                    INPUT := "A/GLR_012_TT03_CHIN",
                    FAULT => "AI_DATA".R12_TT03.Faulty,
                    H_ALM => "AI_DATA".R12_TT03.H_ALM,
                    L_ALM => "AI_DATA".R12_TT03.L_ALM,
                    SCALE_OUT => "AI_DATA".R12_TT03.PV);
   END_IF;
END_REGION

REGION Network 49: ****REACTOR_13****
END_REGION

REGION Network 50: TT01
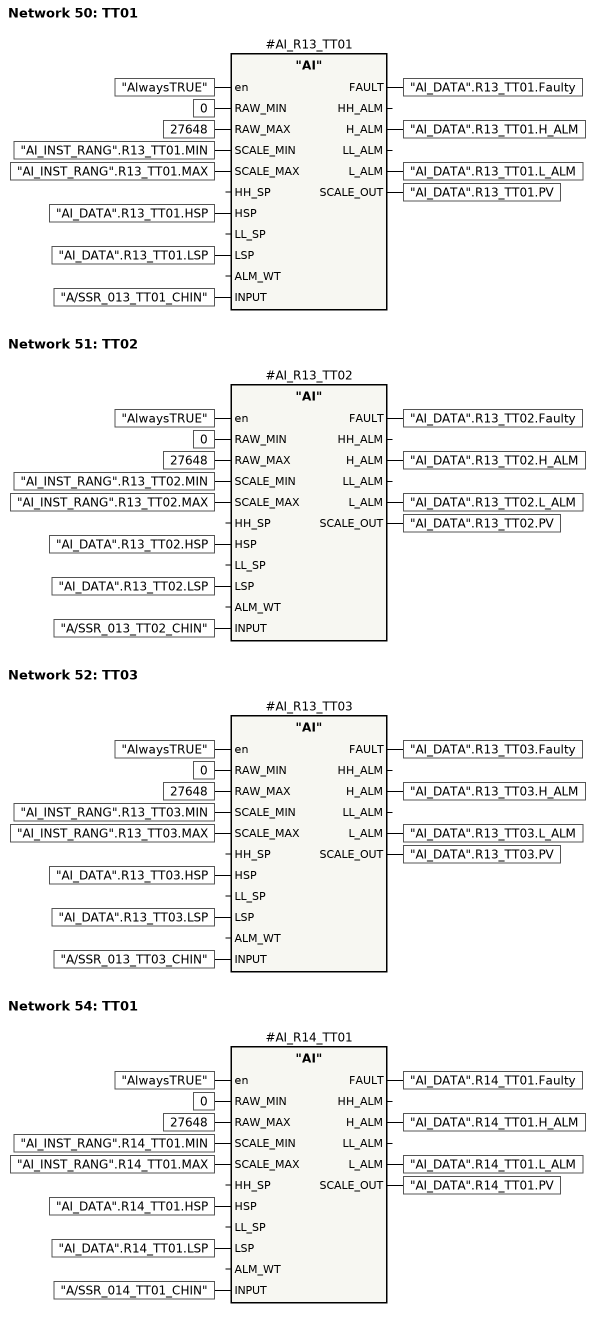
   IF "AlwaysTRUE" THEN
       #AI_R13_TT01(RAW_MIN := 0,   // "AI"
                    RAW_MAX := 27648,
                    SCALE_MIN := "AI_INST_RANG".R13_TT01.MIN,
                    SCALE_MAX := "AI_INST_RANG".R13_TT01.MAX,
                    HSP := "AI_DATA".R13_TT01.HSP,
                    LSP := "AI_DATA".R13_TT01.LSP,
                    INPUT := "A/SSR_013_TT01_CHIN",
                    FAULT => "AI_DATA".R13_TT01.Faulty,
                    H_ALM => "AI_DATA".R13_TT01.H_ALM,
                    L_ALM => "AI_DATA".R13_TT01.L_ALM,
                    SCALE_OUT => "AI_DATA".R13_TT01.PV);
   END_IF;
END_REGION

REGION Network 51: TT02
   IF "AlwaysTRUE" THEN
       #AI_R13_TT02(RAW_MIN := 0,   // "AI"
                    RAW_MAX := 27648,
                    SCALE_MIN := "AI_INST_RANG".R13_TT02.MIN,
                    SCALE_MAX := "AI_INST_RANG".R13_TT02.MAX,
                    HSP := "AI_DATA".R13_TT02.HSP,
                    LSP := "AI_DATA".R13_TT02.LSP,
                    INPUT := "A/SSR_013_TT02_CHIN",
                    FAULT => "AI_DATA".R13_TT02.Faulty,
                    H_ALM => "AI_DATA".R13_TT02.H_ALM,
                    L_ALM => "AI_DATA".R13_TT02.L_ALM,
                    SCALE_OUT => "AI_DATA".R13_TT02.PV);
   END_IF;
END_REGION

REGION Network 52: TT03
   IF "AlwaysTRUE" THEN
       #AI_R13_TT03(RAW_MIN := 0,   // "AI"
                    RAW_MAX := 27648,
                    SCALE_MIN := "AI_INST_RANG".R13_TT03.MIN,
                    SCALE_MAX := "AI_INST_RANG".R13_TT03.MAX,
                    HSP := "AI_DATA".R13_TT03.HSP,
                    LSP := "AI_DATA".R13_TT03.LSP,
                    INPUT := "A/SSR_013_TT03_CHIN",
                    FAULT => "AI_DATA".R13_TT03.Faulty,
                    H_ALM => "AI_DATA".R13_TT03.H_ALM,
                    L_ALM => "AI_DATA".R13_TT03.L_ALM,
                    SCALE_OUT => "AI_DATA".R13_TT03.PV);
   END_IF;
END_REGION

REGION Network 53: ****REACTOR_14****
END_REGION

REGION Network 54: TT01
   IF "AlwaysTRUE" THEN
       #AI_R14_TT01(RAW_MIN := 0,   // "AI"
                    RAW_MAX := 27648,
                    SCALE_MIN := "AI_INST_RANG".R14_TT01.MIN,
                    SCALE_MAX := "AI_INST_RANG".R14_TT01.MAX,
                    HSP := "AI_DATA".R14_TT01.HSP,
                    LSP := "AI_DATA".R14_TT01.LSP,
                    INPUT := "A/SSR_014_TT01_CHIN",
                    FAULT => "AI_DATA".R14_TT01.Faulty,
                    H_ALM => "AI_DATA".R14_TT01.H_ALM,
                    L_ALM => "AI_DATA".R14_TT01.L_ALM,
                    SCALE_OUT => "AI_DATA".R14_TT01.PV);
   END_IF;
END_REGION

REGION Network 55: TT02
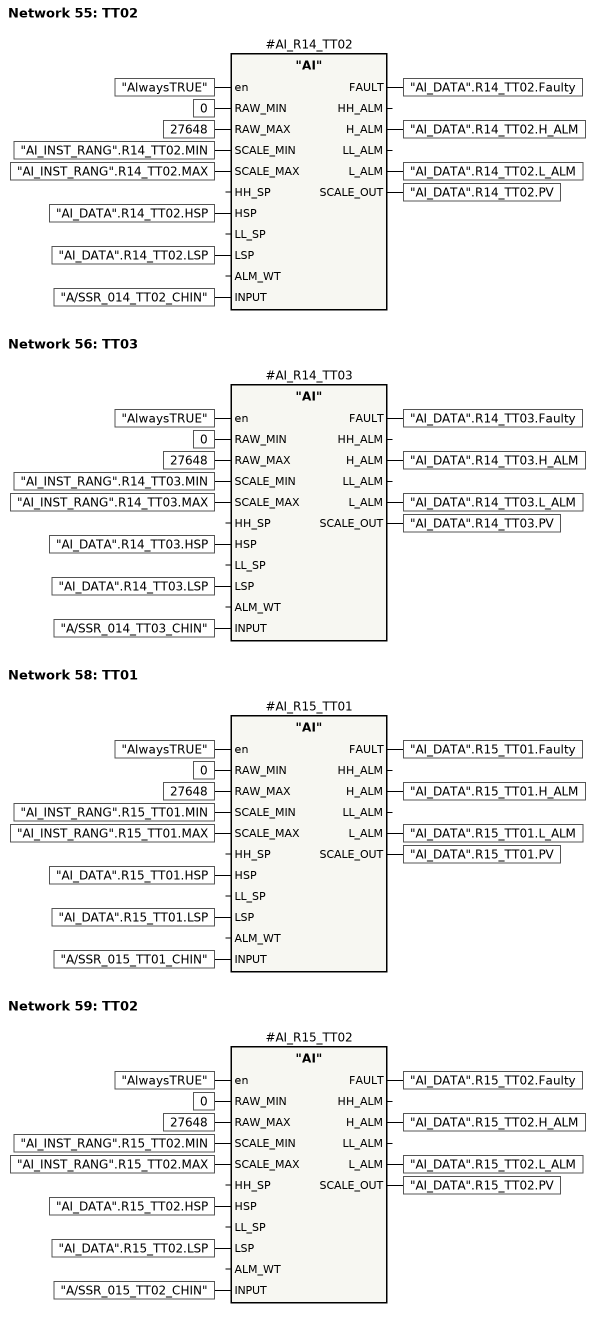
   IF "AlwaysTRUE" THEN
       #AI_R14_TT02(RAW_MIN := 0,   // "AI"
                    RAW_MAX := 27648,
                    SCALE_MIN := "AI_INST_RANG".R14_TT02.MIN,
                    SCALE_MAX := "AI_INST_RANG".R14_TT02.MAX,
                    HSP := "AI_DATA".R14_TT02.HSP,
                    LSP := "AI_DATA".R14_TT02.LSP,
                    INPUT := "A/SSR_014_TT02_CHIN",
                    FAULT => "AI_DATA".R14_TT02.Faulty,
                    H_ALM => "AI_DATA".R14_TT02.H_ALM,
                    L_ALM => "AI_DATA".R14_TT02.L_ALM,
                    SCALE_OUT => "AI_DATA".R14_TT02.PV);
   END_IF;
END_REGION

REGION Network 56: TT03
   IF "AlwaysTRUE" THEN
       #AI_R14_TT03(RAW_MIN := 0,   // "AI"
                    RAW_MAX := 27648,
                    SCALE_MIN := "AI_INST_RANG".R14_TT03.MIN,
                    SCALE_MAX := "AI_INST_RANG".R14_TT03.MAX,
                    HSP := "AI_DATA".R14_TT03.HSP,
                    LSP := "AI_DATA".R14_TT03.LSP,
                    INPUT := "A/SSR_014_TT03_CHIN",
                    FAULT => "AI_DATA".R14_TT03.Faulty,
                    H_ALM => "AI_DATA".R14_TT03.H_ALM,
                    L_ALM => "AI_DATA".R14_TT03.L_ALM,
                    SCALE_OUT => "AI_DATA".R14_TT03.PV);
   END_IF;
END_REGION

REGION Network 57: ****REACTOR_15****
END_REGION

REGION Network 58: TT01
   IF "AlwaysTRUE" THEN
       #AI_R15_TT01(RAW_MIN := 0,   // "AI"
                    RAW_MAX := 27648,
                    SCALE_MIN := "AI_INST_RANG".R15_TT01.MIN,
                    SCALE_MAX := "AI_INST_RANG".R15_TT01.MAX,
                    HSP := "AI_DATA".R15_TT01.HSP,
                    LSP := "AI_DATA".R15_TT01.LSP,
                    INPUT := "A/SSR_015_TT01_CHIN",
                    FAULT => "AI_DATA".R15_TT01.Faulty,
                    H_ALM => "AI_DATA".R15_TT01.H_ALM,
                    L_ALM => "AI_DATA".R15_TT01.L_ALM,
                    SCALE_OUT => "AI_DATA".R15_TT01.PV);
   END_IF;
END_REGION

REGION Network 59: TT02
   IF "AlwaysTRUE" THEN
       #AI_R15_TT02(RAW_MIN := 0,   // "AI"
                    RAW_MAX := 27648,
                    SCALE_MIN := "AI_INST_RANG".R15_TT02.MIN,
                    SCALE_MAX := "AI_INST_RANG".R15_TT02.MAX,
                    HSP := "AI_DATA".R15_TT02.HSP,
                    LSP := "AI_DATA".R15_TT02.LSP,
                    INPUT := "A/SSR_015_TT02_CHIN",
                    FAULT => "AI_DATA".R15_TT02.Faulty,
                    H_ALM => "AI_DATA".R15_TT02.H_ALM,
                    L_ALM => "AI_DATA".R15_TT02.L_ALM,
                    SCALE_OUT => "AI_DATA".R15_TT02.PV);
   END_IF;
END_REGION

REGION Network 60: TT03
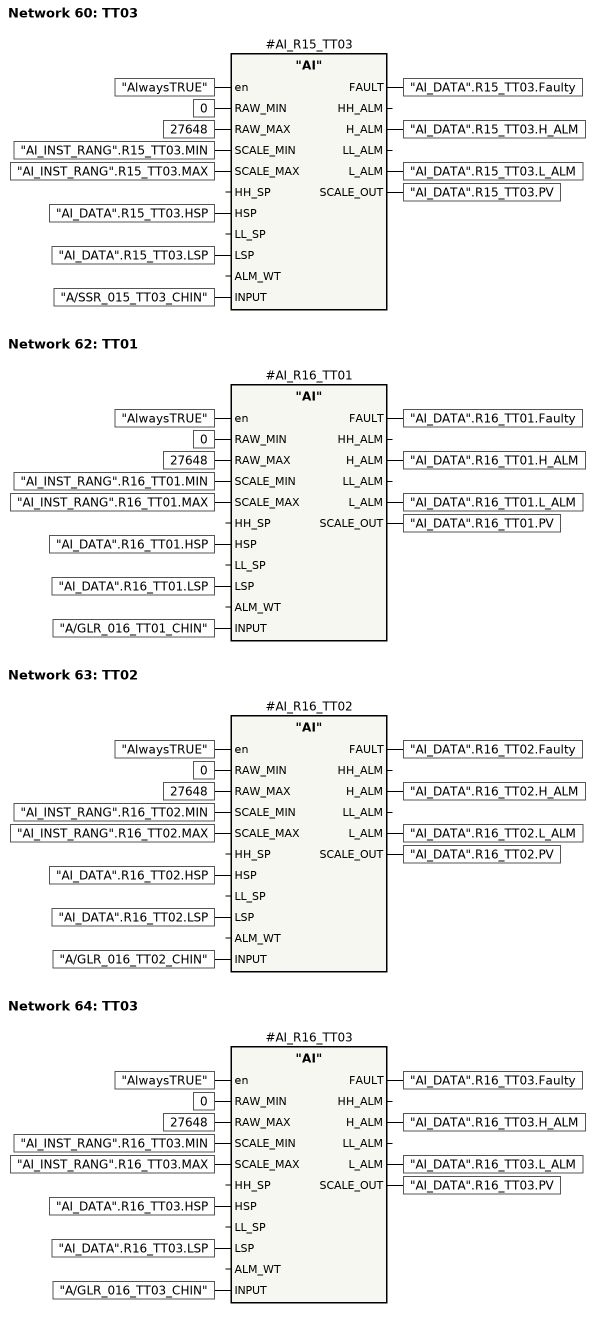
   IF "AlwaysTRUE" THEN
       #AI_R15_TT03(RAW_MIN := 0,   // "AI"
                    RAW_MAX := 27648,
                    SCALE_MIN := "AI_INST_RANG".R15_TT03.MIN,
                    SCALE_MAX := "AI_INST_RANG".R15_TT03.MAX,
                    HSP := "AI_DATA".R15_TT03.HSP,
                    LSP := "AI_DATA".R15_TT03.LSP,
                    INPUT := "A/SSR_015_TT03_CHIN",
                    FAULT => "AI_DATA".R15_TT03.Faulty,
                    H_ALM => "AI_DATA".R15_TT03.H_ALM,
                    L_ALM => "AI_DATA".R15_TT03.L_ALM,
                    SCALE_OUT => "AI_DATA".R15_TT03.PV);
   END_IF;
END_REGION

REGION Network 61: ****REACTOR_16****
END_REGION

REGION Network 62: TT01
   IF "AlwaysTRUE" THEN
       #AI_R16_TT01(RAW_MIN := 0,   // "AI"
                    RAW_MAX := 27648,
                    SCALE_MIN := "AI_INST_RANG".R16_TT01.MIN,
                    SCALE_MAX := "AI_INST_RANG".R16_TT01.MAX,
                    HSP := "AI_DATA".R16_TT01.HSP,
                    LSP := "AI_DATA".R16_TT01.LSP,
                    INPUT := "A/GLR_016_TT01_CHIN",
                    FAULT => "AI_DATA".R16_TT01.Faulty,
                    H_ALM => "AI_DATA".R16_TT01.H_ALM,
                    L_ALM => "AI_DATA".R16_TT01.L_ALM,
                    SCALE_OUT => "AI_DATA".R16_TT01.PV);
   END_IF;
END_REGION

REGION Network 63: TT02
   IF "AlwaysTRUE" THEN
       #AI_R16_TT02(RAW_MIN := 0,   // "AI"
                    RAW_MAX := 27648,
                    SCALE_MIN := "AI_INST_RANG".R16_TT02.MIN,
                    SCALE_MAX := "AI_INST_RANG".R16_TT02.MAX,
                    HSP := "AI_DATA".R16_TT02.HSP,
                    LSP := "AI_DATA".R16_TT02.LSP,
                    INPUT := "A/GLR_016_TT02_CHIN",
                    FAULT => "AI_DATA".R16_TT02.Faulty,
                    H_ALM => "AI_DATA".R16_TT02.H_ALM,
                    L_ALM => "AI_DATA".R16_TT02.L_ALM,
                    SCALE_OUT => "AI_DATA".R16_TT02.PV);
   END_IF;
END_REGION

REGION Network 64: TT03
   IF "AlwaysTRUE" THEN
       #AI_R16_TT03(RAW_MIN := 0,   // "AI"
                    RAW_MAX := 27648,
                    SCALE_MIN := "AI_INST_RANG".R16_TT03.MIN,
                    SCALE_MAX := "AI_INST_RANG".R16_TT03.MAX,
                    HSP := "AI_DATA".R16_TT03.HSP,
                    LSP := "AI_DATA".R16_TT03.LSP,
                    INPUT := "A/GLR_016_TT03_CHIN",
                    FAULT => "AI_DATA".R16_TT03.Faulty,
                    H_ALM => "AI_DATA".R16_TT03.H_ALM,
                    L_ALM => "AI_DATA".R16_TT03.L_ALM,
                    SCALE_OUT => "AI_DATA".R16_TT03.PV);
   END_IF;
END_REGION

REGION Network 65: ****REACTOR_17****
END_REGION

REGION Network 66: TT01
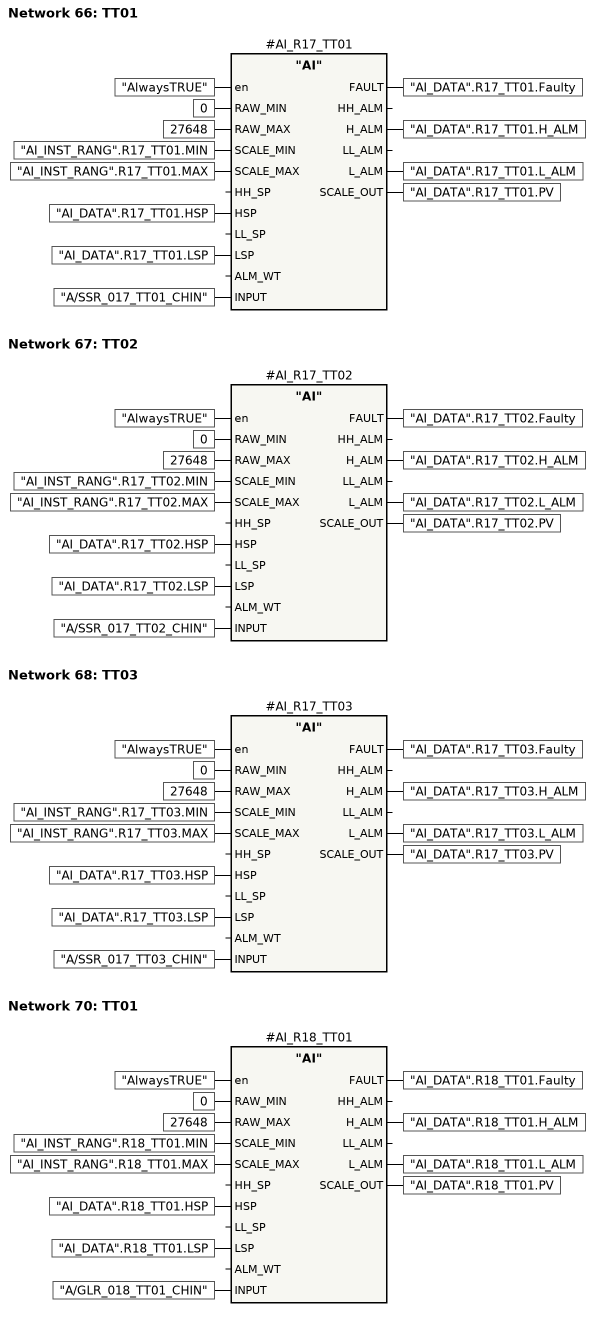
   IF "AlwaysTRUE" THEN
       #AI_R17_TT01(RAW_MIN := 0,   // "AI"
                    RAW_MAX := 27648,
                    SCALE_MIN := "AI_INST_RANG".R17_TT01.MIN,
                    SCALE_MAX := "AI_INST_RANG".R17_TT01.MAX,
                    HSP := "AI_DATA".R17_TT01.HSP,
                    LSP := "AI_DATA".R17_TT01.LSP,
                    INPUT := "A/SSR_017_TT01_CHIN",
                    FAULT => "AI_DATA".R17_TT01.Faulty,
                    H_ALM => "AI_DATA".R17_TT01.H_ALM,
                    L_ALM => "AI_DATA".R17_TT01.L_ALM,
                    SCALE_OUT => "AI_DATA".R17_TT01.PV);
   END_IF;
END_REGION

REGION Network 67: TT02
   IF "AlwaysTRUE" THEN
       #AI_R17_TT02(RAW_MIN := 0,   // "AI"
                    RAW_MAX := 27648,
                    SCALE_MIN := "AI_INST_RANG".R17_TT02.MIN,
                    SCALE_MAX := "AI_INST_RANG".R17_TT02.MAX,
                    HSP := "AI_DATA".R17_TT02.HSP,
                    LSP := "AI_DATA".R17_TT02.LSP,
                    INPUT := "A/SSR_017_TT02_CHIN",
                    FAULT => "AI_DATA".R17_TT02.Faulty,
                    H_ALM => "AI_DATA".R17_TT02.H_ALM,
                    L_ALM => "AI_DATA".R17_TT02.L_ALM,
                    SCALE_OUT => "AI_DATA".R17_TT02.PV);
   END_IF;
END_REGION

REGION Network 68: TT03
   IF "AlwaysTRUE" THEN
       #AI_R17_TT03(RAW_MIN := 0,   // "AI"
                    RAW_MAX := 27648,
                    SCALE_MIN := "AI_INST_RANG".R17_TT03.MIN,
                    SCALE_MAX := "AI_INST_RANG".R17_TT03.MAX,
                    HSP := "AI_DATA".R17_TT03.HSP,
                    LSP := "AI_DATA".R17_TT03.LSP,
                    INPUT := "A/SSR_017_TT03_CHIN",
                    FAULT => "AI_DATA".R17_TT03.Faulty,
                    H_ALM => "AI_DATA".R17_TT03.H_ALM,
                    L_ALM => "AI_DATA".R17_TT03.L_ALM,
                    SCALE_OUT => "AI_DATA".R17_TT03.PV);
   END_IF;
END_REGION

REGION Network 69: ****REACTOR_18****
END_REGION

REGION Network 70: TT01
   IF "AlwaysTRUE" THEN
       #AI_R18_TT01(RAW_MIN := 0,   // "AI"
                    RAW_MAX := 27648,
                    SCALE_MIN := "AI_INST_RANG".R18_TT01.MIN,
                    SCALE_MAX := "AI_INST_RANG".R18_TT01.MAX,
                    HSP := "AI_DATA".R18_TT01.HSP,
                    LSP := "AI_DATA".R18_TT01.LSP,
                    INPUT := "A/GLR_018_TT01_CHIN",
                    FAULT => "AI_DATA".R18_TT01.Faulty,
                    H_ALM => "AI_DATA".R18_TT01.H_ALM,
                    L_ALM => "AI_DATA".R18_TT01.L_ALM,
                    SCALE_OUT => "AI_DATA".R18_TT01.PV);
   END_IF;
END_REGION

REGION Network 71: TT02
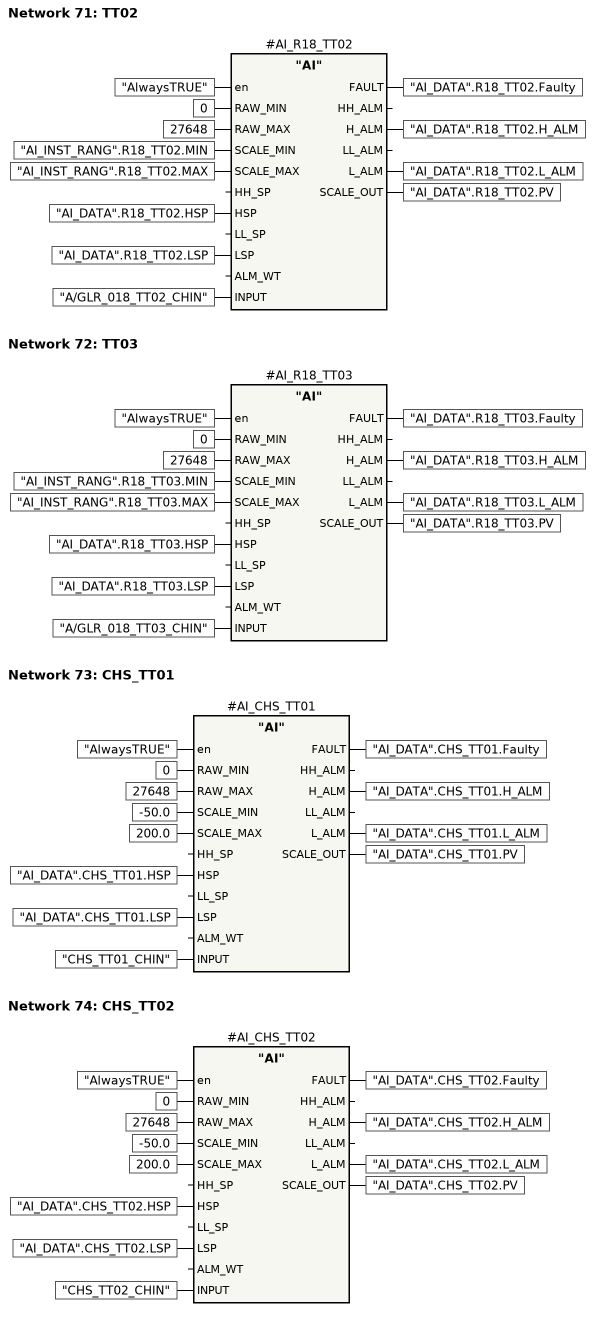
   IF "AlwaysTRUE" THEN
       #AI_R18_TT02(RAW_MIN := 0,   // "AI"
                    RAW_MAX := 27648,
                    SCALE_MIN := "AI_INST_RANG".R18_TT02.MIN,
                    SCALE_MAX := "AI_INST_RANG".R18_TT02.MAX,
                    HSP := "AI_DATA".R18_TT02.HSP,
                    LSP := "AI_DATA".R18_TT02.LSP,
                    INPUT := "A/GLR_018_TT02_CHIN",
                    FAULT => "AI_DATA".R18_TT02.Faulty,
                    H_ALM => "AI_DATA".R18_TT02.H_ALM,
                    L_ALM => "AI_DATA".R18_TT02.L_ALM,
                    SCALE_OUT => "AI_DATA".R18_TT02.PV);
   END_IF;
END_REGION

REGION Network 72: TT03
   IF "AlwaysTRUE" THEN
       #AI_R18_TT03(RAW_MIN := 0,   // "AI"
                    RAW_MAX := 27648,
                    SCALE_MIN := "AI_INST_RANG".R18_TT03.MIN,
                    SCALE_MAX := "AI_INST_RANG".R18_TT03.MAX,
                    HSP := "AI_DATA".R18_TT03.HSP,
                    LSP := "AI_DATA".R18_TT03.LSP,
                    INPUT := "A/GLR_018_TT03_CHIN",
                    FAULT => "AI_DATA".R18_TT03.Faulty,
                    H_ALM => "AI_DATA".R18_TT03.H_ALM,
                    L_ALM => "AI_DATA".R18_TT03.L_ALM,
                    SCALE_OUT => "AI_DATA".R18_TT03.PV);
   END_IF;
END_REGION

REGION Network 73: CHS_TT01
   IF "AlwaysTRUE" THEN
       #AI_CHS_TT01(RAW_MIN := 0,   // "AI"
                    RAW_MAX := 27648,
                    SCALE_MIN := -50.0,
                    SCALE_MAX := 200.0,
                    HSP := "AI_DATA".CHS_TT01.HSP,
                    LSP := "AI_DATA".CHS_TT01.LSP,
                    INPUT := "CHS_TT01_CHIN",
                    FAULT => "AI_DATA".CHS_TT01.Faulty,
                    H_ALM => "AI_DATA".CHS_TT01.H_ALM,
                    L_ALM => "AI_DATA".CHS_TT01.L_ALM,
                    SCALE_OUT => "AI_DATA".CHS_TT01.PV);
   END_IF;
END_REGION

REGION Network 74: CHS_TT02
   IF "AlwaysTRUE" THEN
       #AI_CHS_TT02(RAW_MIN := 0,   // "AI"
                    RAW_MAX := 27648,
                    SCALE_MIN := -50.0,
                    SCALE_MAX := 200.0,
                    HSP := "AI_DATA".CHS_TT02.HSP,
                    LSP := "AI_DATA".CHS_TT02.LSP,
                    INPUT := "CHS_TT02_CHIN",
                    FAULT => "AI_DATA".CHS_TT02.Faulty,
                    H_ALM => "AI_DATA".CHS_TT02.H_ALM,
                    L_ALM => "AI_DATA".CHS_TT02.L_ALM,
                    SCALE_OUT => "AI_DATA".CHS_TT02.PV);
   END_IF;
END_REGION

REGION Network 75: CHS_TT03
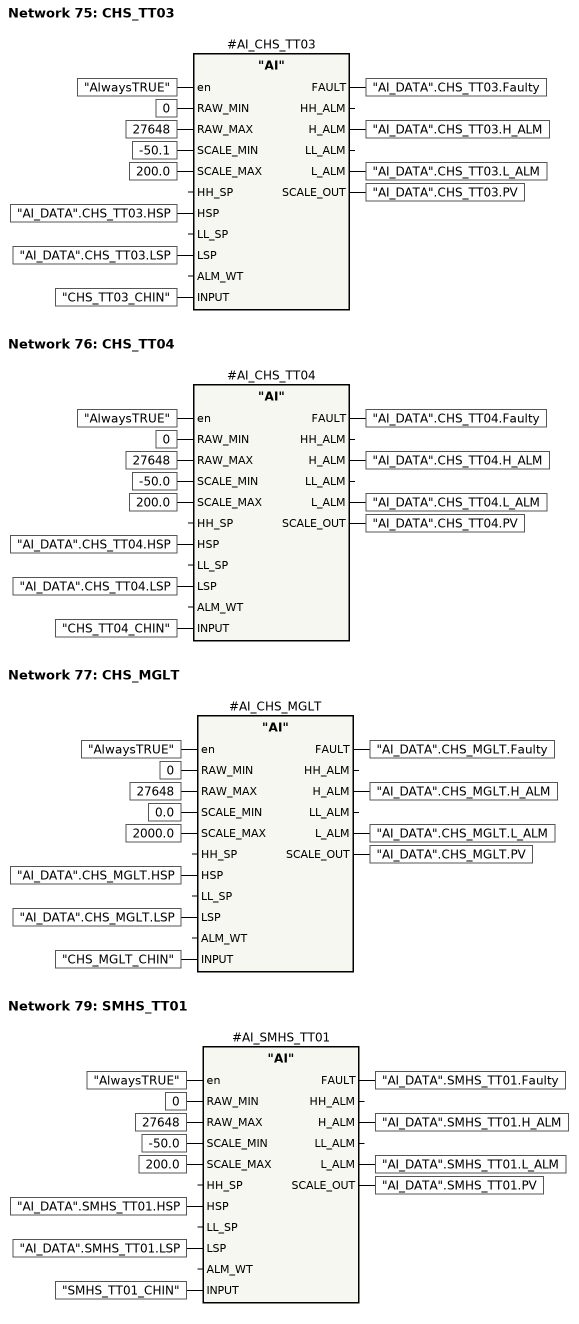
   IF "AlwaysTRUE" THEN
       #AI_CHS_TT03(RAW_MIN := 0,   // "AI"
                    RAW_MAX := 27648,
                    SCALE_MIN := -50.1,
                    SCALE_MAX := 200.0,
                    HSP := "AI_DATA".CHS_TT03.HSP,
                    LSP := "AI_DATA".CHS_TT03.LSP,
                    INPUT := "CHS_TT03_CHIN",
                    FAULT => "AI_DATA".CHS_TT03.Faulty,
                    H_ALM => "AI_DATA".CHS_TT03.H_ALM,
                    L_ALM => "AI_DATA".CHS_TT03.L_ALM,
                    SCALE_OUT => "AI_DATA".CHS_TT03.PV);
   END_IF;
END_REGION

REGION Network 76: CHS_TT04
   IF "AlwaysTRUE" THEN
       #AI_CHS_TT04(RAW_MIN := 0,   // "AI"
                    RAW_MAX := 27648,
                    SCALE_MIN := -50.0,
                    SCALE_MAX := 200.0,
                    HSP := "AI_DATA".CHS_TT04.HSP,
                    LSP := "AI_DATA".CHS_TT04.LSP,
                    INPUT := "CHS_TT04_CHIN",
                    FAULT => "AI_DATA".CHS_TT04.Faulty,
                    H_ALM => "AI_DATA".CHS_TT04.H_ALM,
                    L_ALM => "AI_DATA".CHS_TT04.L_ALM,
                    SCALE_OUT => "AI_DATA".CHS_TT04.PV);
   END_IF;
END_REGION

REGION Network 77: CHS_MGLT
   IF "AlwaysTRUE" THEN
       #AI_CHS_MGLT(RAW_MIN := 0,   // "AI"
                    RAW_MAX := 27648,
                    SCALE_MIN := 0.0,
                    SCALE_MAX := 2000.0,
                    HSP := "AI_DATA".CHS_MGLT.HSP,
                    LSP := "AI_DATA".CHS_MGLT.LSP,
                    INPUT := "CHS_MGLT_CHIN",
                    FAULT => "AI_DATA".CHS_MGLT.Faulty,
                    H_ALM => "AI_DATA".CHS_MGLT.H_ALM,
                    L_ALM => "AI_DATA".CHS_MGLT.L_ALM,
                    SCALE_OUT => "AI_DATA".CHS_MGLT.PV);
   END_IF;
END_REGION

REGION Network 79: SMHS_TT01
   IF "AlwaysTRUE" THEN
       #AI_SMHS_TT01(RAW_MIN := 0,   // "AI"
                     RAW_MAX := 27648,
                     SCALE_MIN := -50.0,
                     SCALE_MAX := 200.0,
                     HSP := "AI_DATA".SMHS_TT01.HSP,
                     LSP := "AI_DATA".SMHS_TT01.LSP,
                     INPUT := "SMHS_TT01_CHIN",
                     FAULT => "AI_DATA".SMHS_TT01.Faulty,
                     H_ALM => "AI_DATA".SMHS_TT01.H_ALM,
                     L_ALM => "AI_DATA".SMHS_TT01.L_ALM,
                     SCALE_OUT => "AI_DATA".SMHS_TT01.PV);
   END_IF;
END_REGION

REGION Network 80: SMCS_TT02
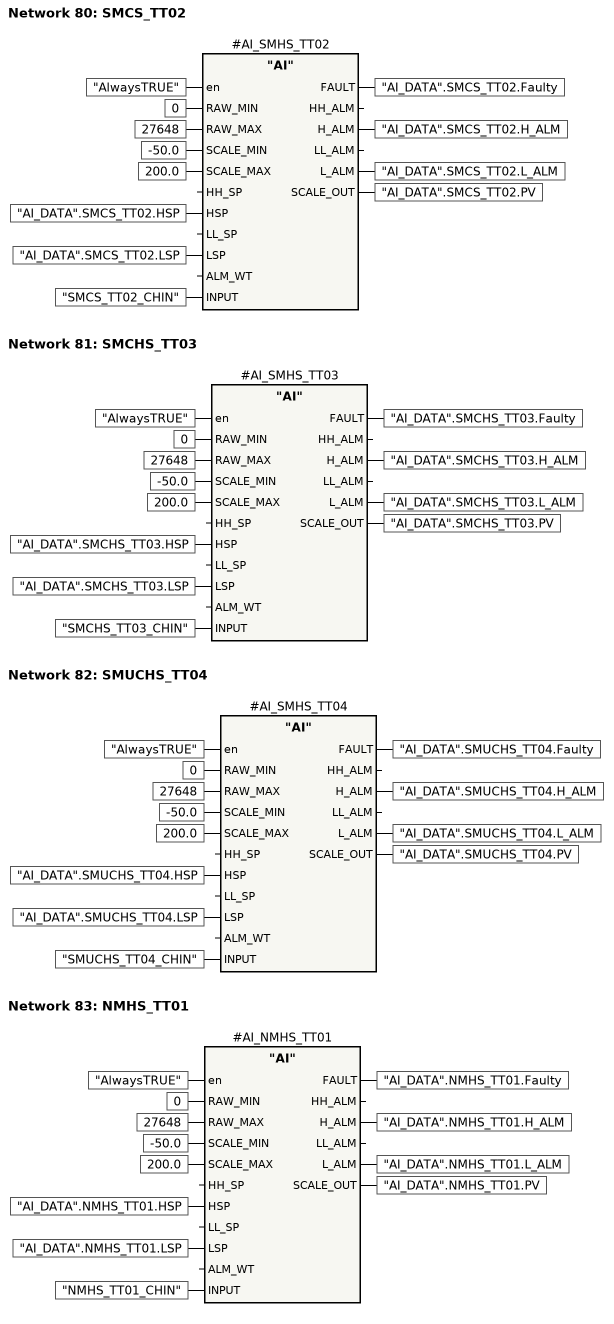
   IF "AlwaysTRUE" THEN
       #AI_SMHS_TT02(RAW_MIN := 0,   // "AI"
                     RAW_MAX := 27648,
                     SCALE_MIN := -50.0,
                     SCALE_MAX := 200.0,
                     HSP := "AI_DATA".SMCS_TT02.HSP,
                     LSP := "AI_DATA".SMCS_TT02.LSP,
                     INPUT := "SMCS_TT02_CHIN",
                     FAULT => "AI_DATA".SMCS_TT02.Faulty,
                     H_ALM => "AI_DATA".SMCS_TT02.H_ALM,
                     L_ALM => "AI_DATA".SMCS_TT02.L_ALM,
                     SCALE_OUT => "AI_DATA".SMCS_TT02.PV);
   END_IF;
END_REGION

REGION Network 81: SMCHS_TT03
   IF "AlwaysTRUE" THEN
       #AI_SMHS_TT03(RAW_MIN := 0,   // "AI"
                     RAW_MAX := 27648,
                     SCALE_MIN := -50.0,
                     SCALE_MAX := 200.0,
                     HSP := "AI_DATA".SMCHS_TT03.HSP,
                     LSP := "AI_DATA".SMCHS_TT03.LSP,
                     INPUT := "SMCHS_TT03_CHIN",
                     FAULT => "AI_DATA".SMCHS_TT03.Faulty,
                     H_ALM => "AI_DATA".SMCHS_TT03.H_ALM,
                     L_ALM => "AI_DATA".SMCHS_TT03.L_ALM,
                     SCALE_OUT => "AI_DATA".SMCHS_TT03.PV);
   END_IF;
END_REGION

REGION Network 82: SMUCHS_TT04
   IF "AlwaysTRUE" THEN
       #AI_SMHS_TT04(RAW_MIN := 0,   // "AI"
                     RAW_MAX := 27648,
                     SCALE_MIN := -50.0,
                     SCALE_MAX := 200.0,
                     HSP := "AI_DATA".SMUCHS_TT04.HSP,
                     LSP := "AI_DATA".SMUCHS_TT04.LSP,
                     INPUT := "SMUCHS_TT04_CHIN",
                     FAULT => "AI_DATA".SMUCHS_TT04.Faulty,
                     H_ALM => "AI_DATA".SMUCHS_TT04.H_ALM,
                     L_ALM => "AI_DATA".SMUCHS_TT04.L_ALM,
                     SCALE_OUT => "AI_DATA".SMUCHS_TT04.PV);
   END_IF;
END_REGION

REGION Network 83: NMHS_TT01
   IF "AlwaysTRUE" THEN
       #AI_NMHS_TT01(RAW_MIN := 0,   // "AI"
                     RAW_MAX := 27648,
                     SCALE_MIN := -50.0,
                     SCALE_MAX := 200.0,
                     HSP := "AI_DATA".NMHS_TT01.HSP,
                     LSP := "AI_DATA".NMHS_TT01.LSP,
                     INPUT := "NMHS_TT01_CHIN",
                     FAULT => "AI_DATA".NMHS_TT01.Faulty,
                     H_ALM => "AI_DATA".NMHS_TT01.H_ALM,
                     L_ALM => "AI_DATA".NMHS_TT01.L_ALM,
                     SCALE_OUT => "AI_DATA".NMHS_TT01.PV);
   END_IF;
END_REGION

REGION Network 84: NMCS_TT02
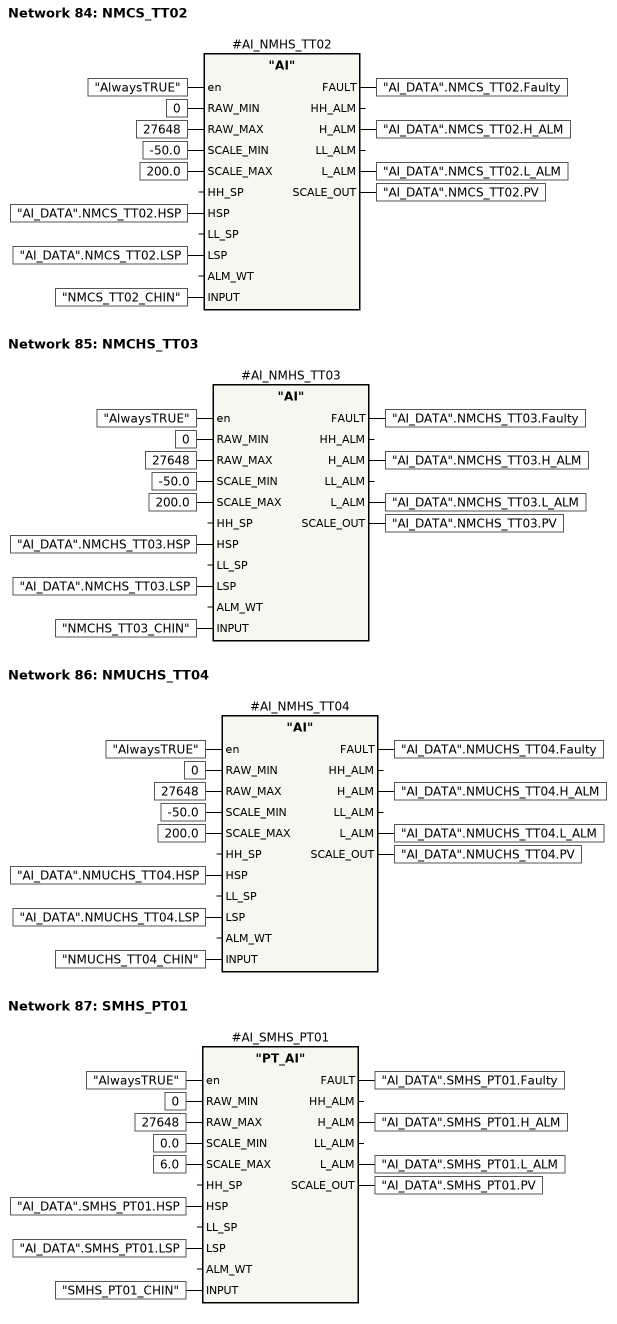
   IF "AlwaysTRUE" THEN
       #AI_NMHS_TT02(RAW_MIN := 0,   // "AI"
                     RAW_MAX := 27648,
                     SCALE_MIN := -50.0,
                     SCALE_MAX := 200.0,
                     HSP := "AI_DATA".NMCS_TT02.HSP,
                     LSP := "AI_DATA".NMCS_TT02.LSP,
                     INPUT := "NMCS_TT02_CHIN",
                     FAULT => "AI_DATA".NMCS_TT02.Faulty,
                     H_ALM => "AI_DATA".NMCS_TT02.H_ALM,
                     L_ALM => "AI_DATA".NMCS_TT02.L_ALM,
                     SCALE_OUT => "AI_DATA".NMCS_TT02.PV);
   END_IF;
END_REGION

REGION Network 85: NMCHS_TT03
   IF "AlwaysTRUE" THEN
       #AI_NMHS_TT03(RAW_MIN := 0,   // "AI"
                     RAW_MAX := 27648,
                     SCALE_MIN := -50.0,
                     SCALE_MAX := 200.0,
                     HSP := "AI_DATA".NMCHS_TT03.HSP,
                     LSP := "AI_DATA".NMCHS_TT03.LSP,
                     INPUT := "NMCHS_TT03_CHIN",
                     FAULT => "AI_DATA".NMCHS_TT03.Faulty,
                     H_ALM => "AI_DATA".NMCHS_TT03.H_ALM,
                     L_ALM => "AI_DATA".NMCHS_TT03.L_ALM,
                     SCALE_OUT => "AI_DATA".NMCHS_TT03.PV);
   END_IF;
END_REGION

REGION Network 86: NMUCHS_TT04
   IF "AlwaysTRUE" THEN
       #AI_NMHS_TT04(RAW_MIN := 0,   // "AI"
                     RAW_MAX := 27648,
                     SCALE_MIN := -50.0,
                     SCALE_MAX := 200.0,
                     HSP := "AI_DATA".NMUCHS_TT04.HSP,
                     LSP := "AI_DATA".NMUCHS_TT04.LSP,
                     INPUT := "NMUCHS_TT04_CHIN",
                     FAULT => "AI_DATA".NMUCHS_TT04.Faulty,
                     H_ALM => "AI_DATA".NMUCHS_TT04.H_ALM,
                     L_ALM => "AI_DATA".NMUCHS_TT04.L_ALM,
                     SCALE_OUT => "AI_DATA".NMUCHS_TT04.PV);
   END_IF;
END_REGION

REGION Network 87: SMHS_PT01
   IF "AlwaysTRUE" THEN
       #AI_SMHS_PT01(RAW_MIN := 0,   // "PT_AI"
                     RAW_MAX := 27648,
                     SCALE_MIN := 0.0,
                     SCALE_MAX := 6.0,
                     HSP := "AI_DATA".SMHS_PT01.HSP,
                     LSP := "AI_DATA".SMHS_PT01.LSP,
                     INPUT := "SMHS_PT01_CHIN",
                     FAULT => "AI_DATA".SMHS_PT01.Faulty,
                     H_ALM => "AI_DATA".SMHS_PT01.H_ALM,
                     L_ALM => "AI_DATA".SMHS_PT01.L_ALM,
                     SCALE_OUT => "AI_DATA".SMHS_PT01.PV);
   END_IF;
END_REGION

REGION Network 88: SMCS_PT02
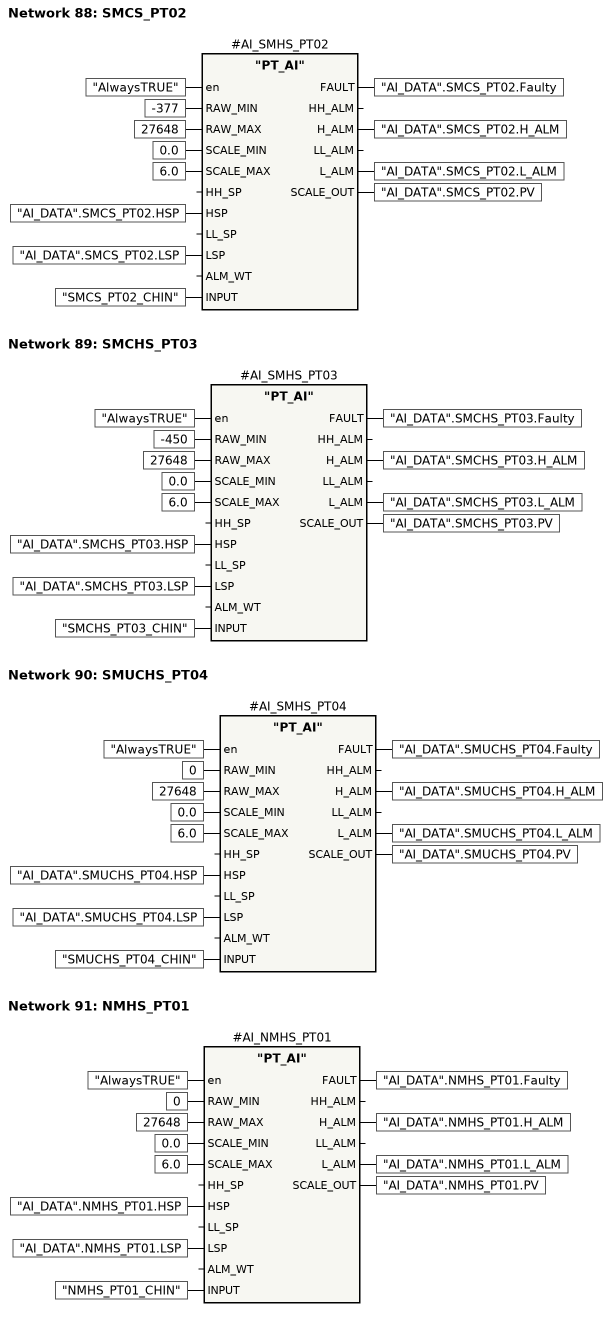
   IF "AlwaysTRUE" THEN
       #AI_SMHS_PT02(RAW_MIN := -377,   // "PT_AI"
                     RAW_MAX := 27648,
                     SCALE_MIN := 0.0,
                     SCALE_MAX := 6.0,
                     HSP := "AI_DATA".SMCS_PT02.HSP,
                     LSP := "AI_DATA".SMCS_PT02.LSP,
                     INPUT := "SMCS_PT02_CHIN",
                     FAULT => "AI_DATA".SMCS_PT02.Faulty,
                     H_ALM => "AI_DATA".SMCS_PT02.H_ALM,
                     L_ALM => "AI_DATA".SMCS_PT02.L_ALM,
                     SCALE_OUT => "AI_DATA".SMCS_PT02.PV);
   END_IF;
END_REGION

REGION Network 89: SMCHS_PT03
   IF "AlwaysTRUE" THEN
       #AI_SMHS_PT03(RAW_MIN := -450,   // "PT_AI"
                     RAW_MAX := 27648,
                     SCALE_MIN := 0.0,
                     SCALE_MAX := 6.0,
                     HSP := "AI_DATA".SMCHS_PT03.HSP,
                     LSP := "AI_DATA".SMCHS_PT03.LSP,
                     INPUT := "SMCHS_PT03_CHIN",
                     FAULT => "AI_DATA".SMCHS_PT03.Faulty,
                     H_ALM => "AI_DATA".SMCHS_PT03.H_ALM,
                     L_ALM => "AI_DATA".SMCHS_PT03.L_ALM,
                     SCALE_OUT => "AI_DATA".SMCHS_PT03.PV);
   END_IF;
END_REGION

REGION Network 90: SMUCHS_PT04
   IF "AlwaysTRUE" THEN
       #AI_SMHS_PT04(RAW_MIN := 0,   // "PT_AI"
                     RAW_MAX := 27648,
                     SCALE_MIN := 0.0,
                     SCALE_MAX := 6.0,
                     HSP := "AI_DATA".SMUCHS_PT04.HSP,
                     LSP := "AI_DATA".SMUCHS_PT04.LSP,
                     INPUT := "SMUCHS_PT04_CHIN",
                     FAULT => "AI_DATA".SMUCHS_PT04.Faulty,
                     H_ALM => "AI_DATA".SMUCHS_PT04.H_ALM,
                     L_ALM => "AI_DATA".SMUCHS_PT04.L_ALM,
                     SCALE_OUT => "AI_DATA".SMUCHS_PT04.PV);
   END_IF;
END_REGION

REGION Network 91: NMHS_PT01
   IF "AlwaysTRUE" THEN
       #AI_NMHS_PT01(RAW_MIN := 0,   // "PT_AI"
                     RAW_MAX := 27648,
                     SCALE_MIN := 0.0,
                     SCALE_MAX := 6.0,
                     HSP := "AI_DATA".NMHS_PT01.HSP,
                     LSP := "AI_DATA".NMHS_PT01.LSP,
                     INPUT := "NMHS_PT01_CHIN",
                     FAULT => "AI_DATA".NMHS_PT01.Faulty,
                     H_ALM => "AI_DATA".NMHS_PT01.H_ALM,
                     L_ALM => "AI_DATA".NMHS_PT01.L_ALM,
                     SCALE_OUT => "AI_DATA".NMHS_PT01.PV);
   END_IF;
END_REGION

REGION Network 92: NMHS_PT02
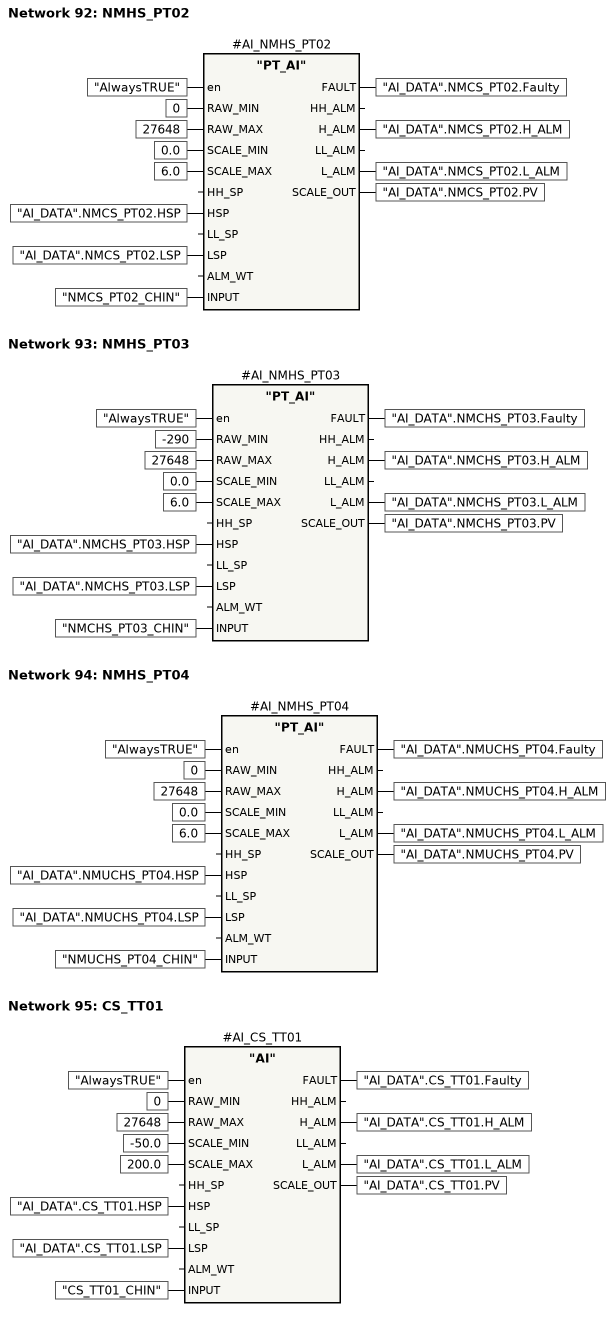
   IF "AlwaysTRUE" THEN
       #AI_NMHS_PT02(RAW_MIN := 0,   // "PT_AI"
                     RAW_MAX := 27648,
                     SCALE_MIN := 0.0,
                     SCALE_MAX := 6.0,
                     HSP := "AI_DATA".NMCS_PT02.HSP,
                     LSP := "AI_DATA".NMCS_PT02.LSP,
                     INPUT := "NMCS_PT02_CHIN",
                     FAULT => "AI_DATA".NMCS_PT02.Faulty,
                     H_ALM => "AI_DATA".NMCS_PT02.H_ALM,
                     L_ALM => "AI_DATA".NMCS_PT02.L_ALM,
                     SCALE_OUT => "AI_DATA".NMCS_PT02.PV);
   END_IF;
END_REGION

REGION Network 93: NMHS_PT03
   IF "AlwaysTRUE" THEN
       #AI_NMHS_PT03(RAW_MIN := -290,   // "PT_AI"
                     RAW_MAX := 27648,
                     SCALE_MIN := 0.0,
                     SCALE_MAX := 6.0,
                     HSP := "AI_DATA".NMCHS_PT03.HSP,
                     LSP := "AI_DATA".NMCHS_PT03.LSP,
                     INPUT := "NMCHS_PT03_CHIN",
                     FAULT => "AI_DATA".NMCHS_PT03.Faulty,
                     H_ALM => "AI_DATA".NMCHS_PT03.H_ALM,
                     L_ALM => "AI_DATA".NMCHS_PT03.L_ALM,
                     SCALE_OUT => "AI_DATA".NMCHS_PT03.PV);
   END_IF;
END_REGION

REGION Network 94: NMHS_PT04
   IF "AlwaysTRUE" THEN
       #AI_NMHS_PT04(RAW_MIN := 0,   // "PT_AI"
                     RAW_MAX := 27648,
                     SCALE_MIN := 0.0,
                     SCALE_MAX := 6.0,
                     HSP := "AI_DATA".NMUCHS_PT04.HSP,
                     LSP := "AI_DATA".NMUCHS_PT04.LSP,
                     INPUT := "NMUCHS_PT04_CHIN",
                     FAULT => "AI_DATA".NMUCHS_PT04.Faulty,
                     H_ALM => "AI_DATA".NMUCHS_PT04.H_ALM,
                     L_ALM => "AI_DATA".NMUCHS_PT04.L_ALM,
                     SCALE_OUT => "AI_DATA".NMUCHS_PT04.PV);
   END_IF;
END_REGION

REGION Network 95: CS_TT01
   IF "AlwaysTRUE" THEN
       #AI_CS_TT01(RAW_MIN := 0,   // "AI"
                   RAW_MAX := 27648,
                   SCALE_MIN := -50.0,
                   SCALE_MAX := 200.0,
                   HSP := "AI_DATA".CS_TT01.HSP,
                   LSP := "AI_DATA".CS_TT01.LSP,
                   INPUT := "CS_TT01_CHIN",
                   FAULT => "AI_DATA".CS_TT01.Faulty,
                   H_ALM => "AI_DATA".CS_TT01.H_ALM,
                   L_ALM => "AI_DATA".CS_TT01.L_ALM,
                   SCALE_OUT => "AI_DATA".CS_TT01.PV);
   END_IF;
END_REGION

REGION Network 96: CS_TT02
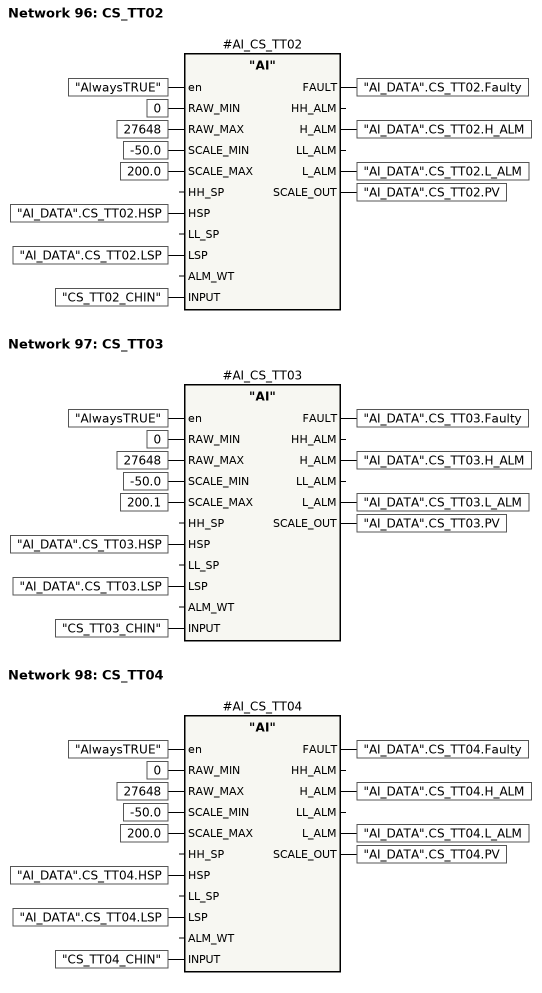
   IF "AlwaysTRUE" THEN
       #AI_CS_TT02(RAW_MIN := 0,   // "AI"
                   RAW_MAX := 27648,
                   SCALE_MIN := -50.0,
                   SCALE_MAX := 200.0,
                   HSP := "AI_DATA".CS_TT02.HSP,
                   LSP := "AI_DATA".CS_TT02.LSP,
                   INPUT := "CS_TT02_CHIN",
                   FAULT => "AI_DATA".CS_TT02.Faulty,
                   H_ALM => "AI_DATA".CS_TT02.H_ALM,
                   L_ALM => "AI_DATA".CS_TT02.L_ALM,
                   SCALE_OUT => "AI_DATA".CS_TT02.PV);
   END_IF;
END_REGION

REGION Network 97: CS_TT03
   IF "AlwaysTRUE" THEN
       #AI_CS_TT03(RAW_MIN := 0,   // "AI"
                   RAW_MAX := 27648,
                   SCALE_MIN := -50.0,
                   SCALE_MAX := 200.1,
                   HSP := "AI_DATA".CS_TT03.HSP,
                   LSP := "AI_DATA".CS_TT03.LSP,
                   INPUT := "CS_TT03_CHIN",
                   FAULT => "AI_DATA".CS_TT03.Faulty,
                   H_ALM => "AI_DATA".CS_TT03.H_ALM,
                   L_ALM => "AI_DATA".CS_TT03.L_ALM,
                   SCALE_OUT => "AI_DATA".CS_TT03.PV);
   END_IF;
END_REGION

REGION Network 98: CS_TT04
   IF "AlwaysTRUE" THEN
       #AI_CS_TT04(RAW_MIN := 0,   // "AI"
                   RAW_MAX := 27648,
                   SCALE_MIN := -50.0,
                   SCALE_MAX := 200.0,
                   HSP := "AI_DATA".CS_TT04.HSP,
                   LSP := "AI_DATA".CS_TT04.LSP,
                   INPUT := "CS_TT04_CHIN",
                   FAULT => "AI_DATA".CS_TT04.Faulty,
                   H_ALM => "AI_DATA".CS_TT04.H_ALM,
                   L_ALM => "AI_DATA".CS_TT04.L_ALM,
                   SCALE_OUT => "AI_DATA".CS_TT04.PV);
   END_IF;
END_REGION

REGION Network 99: CS_MGLT
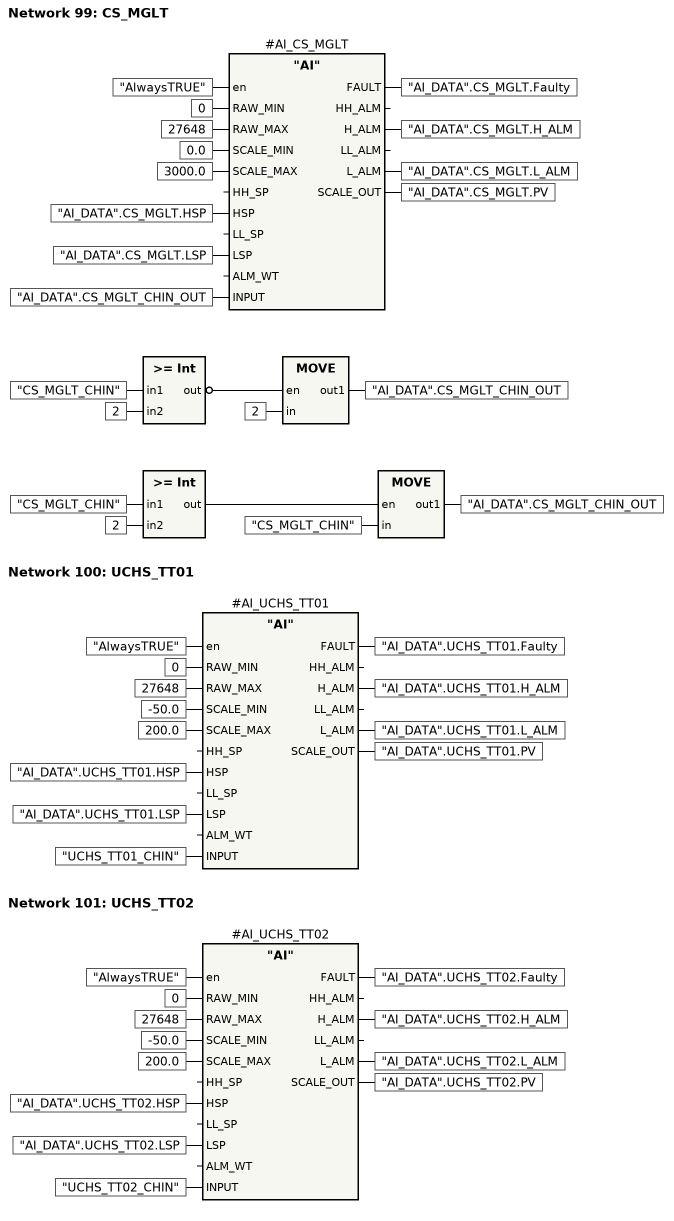
   IF "AlwaysTRUE" THEN
       #AI_CS_MGLT(RAW_MIN := 0,   // "AI"
                   RAW_MAX := 27648,
                   SCALE_MIN := 0.0,
                   SCALE_MAX := 3000.0,
                   HSP := "AI_DATA".CS_MGLT.HSP,
                   LSP := "AI_DATA".CS_MGLT.LSP,
                   INPUT := "AI_DATA".CS_MGLT_CHIN_OUT,
                   FAULT => "AI_DATA".CS_MGLT.Faulty,
                   H_ALM => "AI_DATA".CS_MGLT.H_ALM,
                   L_ALM => "AI_DATA".CS_MGLT.L_ALM,
                   SCALE_OUT => "AI_DATA".CS_MGLT.PV);
   END_IF;
   IF NOT ("CS_MGLT_CHIN" >= 2) THEN "AI_DATA".CS_MGLT_CHIN_OUT := 2; END_IF;
   IF "CS_MGLT_CHIN" >= 2 THEN "AI_DATA".CS_MGLT_CHIN_OUT := "CS_MGLT_CHIN"; END_IF;
END_REGION

REGION Network 100: UCHS_TT01
   IF "AlwaysTRUE" THEN
       #AI_UCHS_TT01(RAW_MIN := 0,   // "AI"
                     RAW_MAX := 27648,
                     SCALE_MIN := -50.0,
                     SCALE_MAX := 200.0,
                     HSP := "AI_DATA".UCHS_TT01.HSP,
                     LSP := "AI_DATA".UCHS_TT01.LSP,
                     INPUT := "UCHS_TT01_CHIN",
                     FAULT => "AI_DATA".UCHS_TT01.Faulty,
                     H_ALM => "AI_DATA".UCHS_TT01.H_ALM,
                     L_ALM => "AI_DATA".UCHS_TT01.L_ALM,
                     SCALE_OUT => "AI_DATA".UCHS_TT01.PV);
   END_IF;
END_REGION

REGION Network 101: UCHS_TT02
   IF "AlwaysTRUE" THEN
       #AI_UCHS_TT02(RAW_MIN := 0,   // "AI"
                     RAW_MAX := 27648,
                     SCALE_MIN := -50.0,
                     SCALE_MAX := 200.0,
                     HSP := "AI_DATA".UCHS_TT02.HSP,
                     LSP := "AI_DATA".UCHS_TT02.LSP,
                     INPUT := "UCHS_TT02_CHIN",
                     FAULT => "AI_DATA".UCHS_TT02.Faulty,
                     H_ALM => "AI_DATA".UCHS_TT02.H_ALM,
                     L_ALM => "AI_DATA".UCHS_TT02.L_ALM,
                     SCALE_OUT => "AI_DATA".UCHS_TT02.PV);
   END_IF;
END_REGION

REGION Network 102: UCHS_TT03
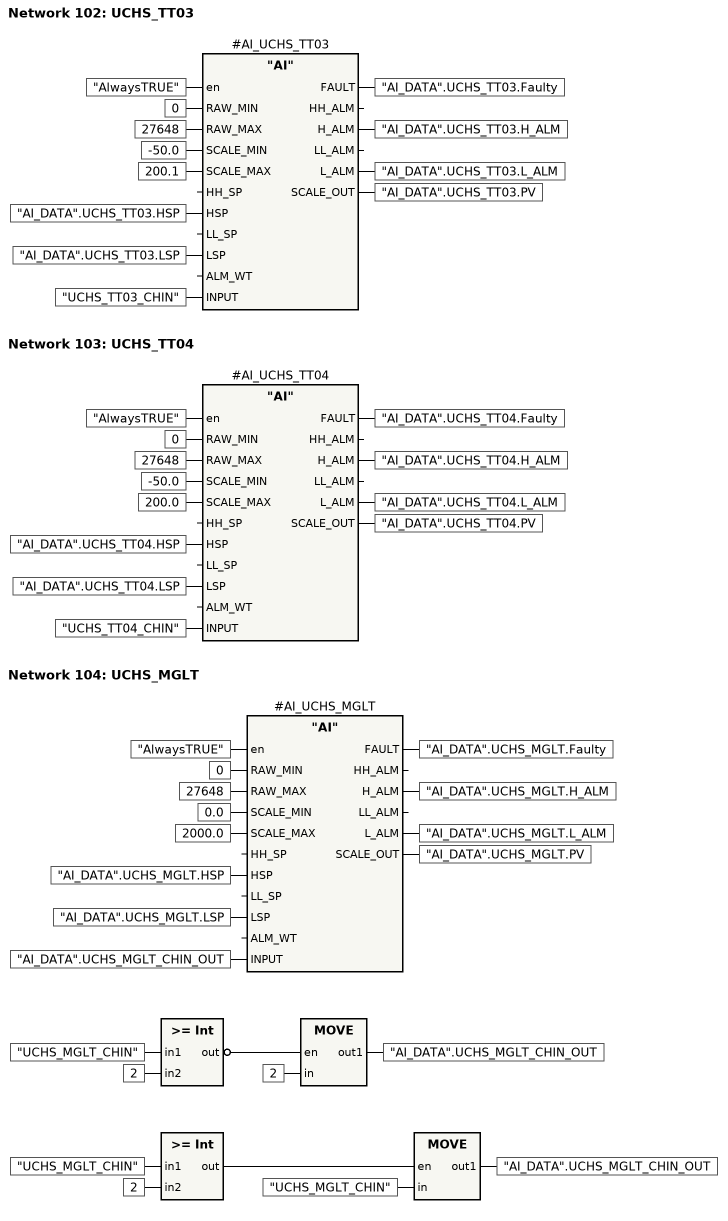
   IF "AlwaysTRUE" THEN
       #AI_UCHS_TT03(RAW_MIN := 0,   // "AI"
                     RAW_MAX := 27648,
                     SCALE_MIN := -50.0,
                     SCALE_MAX := 200.1,
                     HSP := "AI_DATA".UCHS_TT03.HSP,
                     LSP := "AI_DATA".UCHS_TT03.LSP,
                     INPUT := "UCHS_TT03_CHIN",
                     FAULT => "AI_DATA".UCHS_TT03.Faulty,
                     H_ALM => "AI_DATA".UCHS_TT03.H_ALM,
                     L_ALM => "AI_DATA".UCHS_TT03.L_ALM,
                     SCALE_OUT => "AI_DATA".UCHS_TT03.PV);
   END_IF;
END_REGION

REGION Network 103: UCHS_TT04
   IF "AlwaysTRUE" THEN
       #AI_UCHS_TT04(RAW_MIN := 0,   // "AI"
                     RAW_MAX := 27648,
                     SCALE_MIN := -50.0,
                     SCALE_MAX := 200.0,
                     HSP := "AI_DATA".UCHS_TT04.HSP,
                     LSP := "AI_DATA".UCHS_TT04.LSP,
                     INPUT := "UCHS_TT04_CHIN",
                     FAULT => "AI_DATA".UCHS_TT04.Faulty,
                     H_ALM => "AI_DATA".UCHS_TT04.H_ALM,
                     L_ALM => "AI_DATA".UCHS_TT04.L_ALM,
                     SCALE_OUT => "AI_DATA".UCHS_TT04.PV);
   END_IF;
END_REGION

REGION Network 104: UCHS_MGLT
   IF "AlwaysTRUE" THEN
       #AI_UCHS_MGLT(RAW_MIN := 0,   // "AI"
                     RAW_MAX := 27648,
                     SCALE_MIN := 0.0,
                     SCALE_MAX := 2000.0,
                     HSP := "AI_DATA".UCHS_MGLT.HSP,
                     LSP := "AI_DATA".UCHS_MGLT.LSP,
                     INPUT := "AI_DATA".UCHS_MGLT_CHIN_OUT,
                     FAULT => "AI_DATA".UCHS_MGLT.Faulty,
                     H_ALM => "AI_DATA".UCHS_MGLT.H_ALM,
                     L_ALM => "AI_DATA".UCHS_MGLT.L_ALM,
                     SCALE_OUT => "AI_DATA".UCHS_MGLT.PV);
   END_IF;
   IF NOT ("UCHS_MGLT_CHIN" >= 2) THEN "AI_DATA".UCHS_MGLT_CHIN_OUT := 2; END_IF;
   IF "UCHS_MGLT_CHIN" >= 2 THEN "AI_DATA".UCHS_MGLT_CHIN_OUT := "UCHS_MGLT_CHIN"; END_IF;
END_REGION

REGION Network 105: HS_TT01
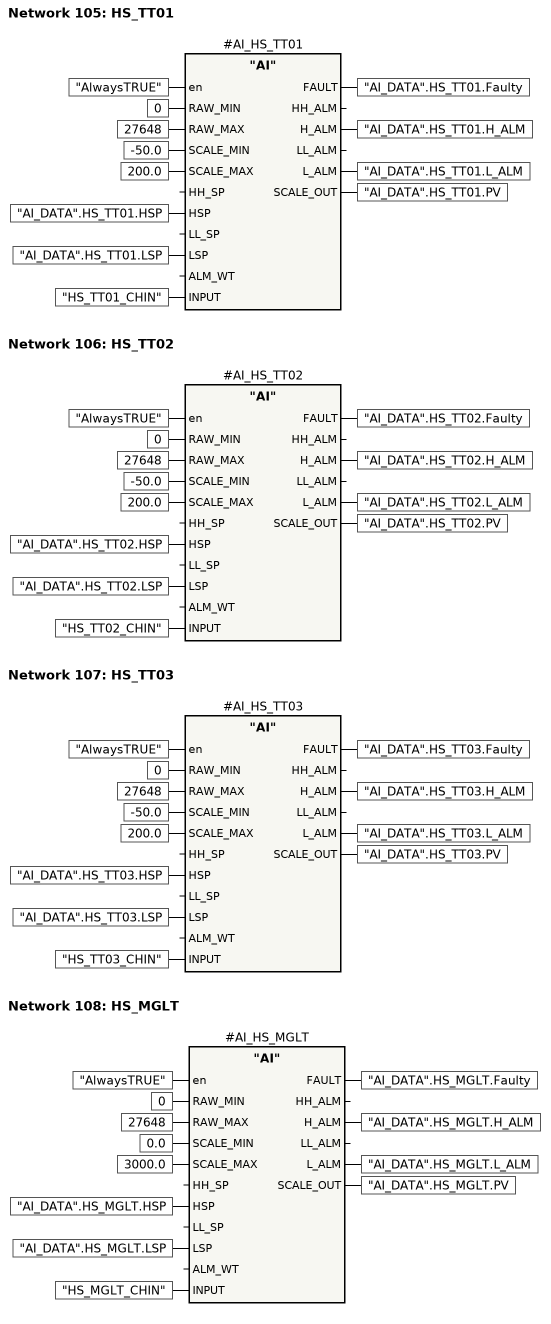
   IF "AlwaysTRUE" THEN
       #AI_HS_TT01(RAW_MIN := 0,   // "AI"
                   RAW_MAX := 27648,
                   SCALE_MIN := -50.0,
                   SCALE_MAX := 200.0,
                   HSP := "AI_DATA".HS_TT01.HSP,
                   LSP := "AI_DATA".HS_TT01.LSP,
                   INPUT := "HS_TT01_CHIN",
                   FAULT => "AI_DATA".HS_TT01.Faulty,
                   H_ALM => "AI_DATA".HS_TT01.H_ALM,
                   L_ALM => "AI_DATA".HS_TT01.L_ALM,
                   SCALE_OUT => "AI_DATA".HS_TT01.PV);
   END_IF;
END_REGION

REGION Network 106: HS_TT02
   IF "AlwaysTRUE" THEN
       #AI_HS_TT02(RAW_MIN := 0,   // "AI"
                   RAW_MAX := 27648,
                   SCALE_MIN := -50.0,
                   SCALE_MAX := 200.0,
                   HSP := "AI_DATA".HS_TT02.HSP,
                   LSP := "AI_DATA".HS_TT02.LSP,
                   INPUT := "HS_TT02_CHIN",
                   FAULT => "AI_DATA".HS_TT02.Faulty,
                   H_ALM => "AI_DATA".HS_TT02.H_ALM,
                   L_ALM => "AI_DATA".HS_TT02.L_ALM,
                   SCALE_OUT => "AI_DATA".HS_TT02.PV);
   END_IF;
END_REGION

REGION Network 107: HS_TT03
   IF "AlwaysTRUE" THEN
       #AI_HS_TT03(RAW_MIN := 0,   // "AI"
                   RAW_MAX := 27648,
                   SCALE_MIN := -50.0,
                   SCALE_MAX := 200.0,
                   HSP := "AI_DATA".HS_TT03.HSP,
                   LSP := "AI_DATA".HS_TT03.LSP,
                   INPUT := "HS_TT03_CHIN",
                   FAULT => "AI_DATA".HS_TT03.Faulty,
                   H_ALM => "AI_DATA".HS_TT03.H_ALM,
                   L_ALM => "AI_DATA".HS_TT03.L_ALM,
                   SCALE_OUT => "AI_DATA".HS_TT03.PV);
   END_IF;
END_REGION

REGION Network 108: HS_MGLT
   IF "AlwaysTRUE" THEN
       #AI_HS_MGLT(RAW_MIN := 0,   // "AI"
                   RAW_MAX := 27648,
                   SCALE_MIN := 0.0,
                   SCALE_MAX := 3000.0,
                   HSP := "AI_DATA".HS_MGLT.HSP,
                   LSP := "AI_DATA".HS_MGLT.LSP,
                   INPUT := "HS_MGLT_CHIN",
                   FAULT => "AI_DATA".HS_MGLT.Faulty,
                   H_ALM => "AI_DATA".HS_MGLT.H_ALM,
                   L_ALM => "AI_DATA".HS_MGLT.L_ALM,
                   SCALE_OUT => "AI_DATA".HS_MGLT.PV);
   END_IF;
END_REGION

REGION Network 110: SCRB_001_PH01
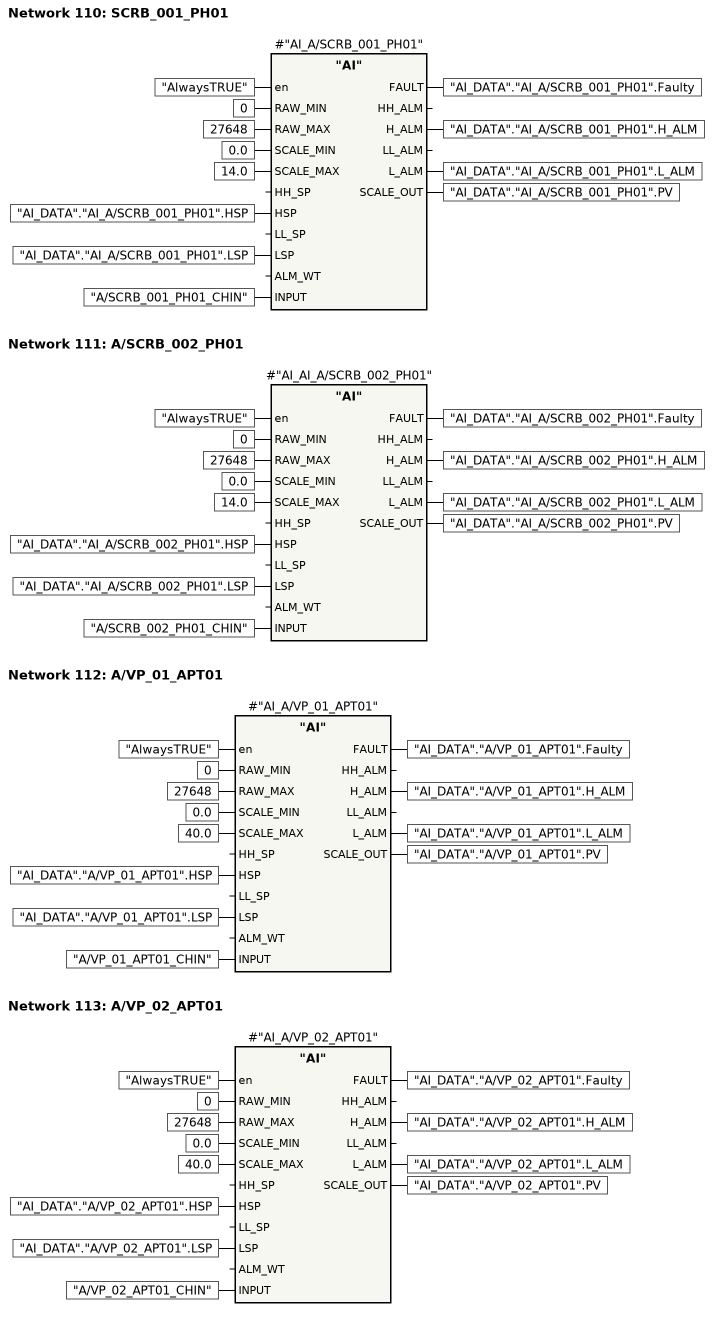
   IF "AlwaysTRUE" THEN
       #"AI_A/SCRB_001_PH01"(RAW_MIN := 0,   // "AI"
                             RAW_MAX := 27648,
                             SCALE_MIN := 0.0,
                             SCALE_MAX := 14.0,
                             HSP := "AI_DATA"."AI_A/SCRB_001_PH01".HSP,
                             LSP := "AI_DATA"."AI_A/SCRB_001_PH01".LSP,
                             INPUT := "A/SCRB_001_PH01_CHIN",
                             FAULT => "AI_DATA"."AI_A/SCRB_001_PH01".Faulty,
                             H_ALM => "AI_DATA"."AI_A/SCRB_001_PH01".H_ALM,
                             L_ALM => "AI_DATA"."AI_A/SCRB_001_PH01".L_ALM,
                             SCALE_OUT => "AI_DATA"."AI_A/SCRB_001_PH01".PV);
   END_IF;
END_REGION

REGION Network 111: A/SCRB_002_PH01
   IF "AlwaysTRUE" THEN
       #"AI_AI_A/SCRB_002_PH01"(RAW_MIN := 0,   // "AI"
                               RAW_MAX := 27648,
                               SCALE_MIN := 0.0,
                               SCALE_MAX := 14.0,
                               HSP := "AI_DATA"."AI_A/SCRB_002_PH01".HSP,
                               LSP := "AI_DATA"."AI_A/SCRB_002_PH01".LSP,
                               INPUT := "A/SCRB_002_PH01_CHIN",
                               FAULT => "AI_DATA"."AI_A/SCRB_002_PH01".Faulty,
                               H_ALM => "AI_DATA"."AI_A/SCRB_002_PH01".H_ALM,
                               L_ALM => "AI_DATA"."AI_A/SCRB_002_PH01".L_ALM,
                               SCALE_OUT => "AI_DATA"."AI_A/SCRB_002_PH01".PV);
   END_IF;
END_REGION

REGION Network 112: A/VP_01_APT01
   IF "AlwaysTRUE" THEN
       #"AI_A/VP_01_APT01"(RAW_MIN := 0,   // "AI"
                           RAW_MAX := 27648,
                           SCALE_MIN := 0.0,
                           SCALE_MAX := 40.0,
                           HSP := "AI_DATA"."A/VP_01_APT01".HSP,
                           LSP := "AI_DATA"."A/VP_01_APT01".LSP,
                           INPUT := "A/VP_01_APT01_CHIN",
                           FAULT => "AI_DATA"."A/VP_01_APT01".Faulty,
                           H_ALM => "AI_DATA"."A/VP_01_APT01".H_ALM,
                           L_ALM => "AI_DATA"."A/VP_01_APT01".L_ALM,
                           SCALE_OUT => "AI_DATA"."A/VP_01_APT01".PV);
   END_IF;
END_REGION

REGION Network 113: A/VP_02_APT01
   IF "AlwaysTRUE" THEN
       #"AI_A/VP_02_APT01"(RAW_MIN := 0,   // "AI"
                           RAW_MAX := 27648,
                           SCALE_MIN := 0.0,
                           SCALE_MAX := 40.0,
                           HSP := "AI_DATA"."A/VP_02_APT01".HSP,
                           LSP := "AI_DATA"."A/VP_02_APT01".LSP,
                           INPUT := "A/VP_02_APT01_CHIN",
                           FAULT => "AI_DATA"."A/VP_02_APT01".Faulty,
                           H_ALM => "AI_DATA"."A/VP_02_APT01".H_ALM,
                           L_ALM => "AI_DATA"."A/VP_02_APT01".L_ALM,
                           SCALE_OUT => "AI_DATA"."A/VP_02_APT01".PV);
   END_IF;
END_REGION

REGION Network 114: A/ANFD_001_APT01
